  rq_init_comm_if_connected(9, "1")
  rq_init_comm_if_connected(2, "2")
  rq_init_comm_if_connected(3, "3")
  rq_init_comm_if_connected(4, "4")
  rq_print_connected_grippers()
  rq_gripper_communication_thread = run rq_gripper_communication()
  set_closed_norm(97.6470588235294, 1)
  set_open_norm(1.1764705882352942, 1)
  set_closed_mm(0.0, 1)
  set_open_mm(53.0, 1)
  set_closed_norm(100.0, 2)
  set_open_norm(0.0, 2)
  set_closed_mm(0.0, 2)
  set_open_mm(50.0, 2)
  set_closed_norm(100.0, 3)
  set_open_norm(0.0, 3)
  set_closed_mm(0.0, 3)
  set_open_mm(50.0, 3)
  set_closed_norm(100.0, 4)
  set_open_norm(0.0, 4)
  set_closed_mm(0.0, 4)
  set_open_mm(50.0, 4)
  rq_current_limit_enabled = False
  while(not rq_gripper_communication_thread_started):
      sync()
  end
  # end: URCap Installation Node
  global AMR_Position=struct(position_identifier=0, x1=0, x2=0, y1=0, y2=0, theta1=0, theta2=0)
  global CAM_Pose=p[0,0,0,0,0,0]
  global CAM_Relation=""
  global CMD_Abort=  False
  global CMD_Clear=  False
  global CMD_Reset=  False
  global CMD_Start=  False
  global CMD_Suspend=  False
  global CMD_Unhold=  False
  global CMD_Unsuspend=  False
  global CNT_Rack_Output=0
  global FNC_Freedrive=  False
  global PRC_TubCounter=0
  global PRC_TubNumber=0
  global STP=0
  global easyPickCount=0
  global easyPickCount_1=0
  global easyPickCount_2=0
  global easyPickCount_3=0
  global easyPickNoObj=0
  global easyPickNoObj_1=0
  global easyPickNoObj_2=0
  global easyPickNoObj_3=0
  global easyPickParts=0
  global easyPickParts_1=0
  global easyPickParts_2=0
  global easyPickParts_3=0
  global TMR_Barcode=0
  global Waypoint_6_p=p[.008800512419, -.547926542621, .402696567415, -.589884378425, -.007228654778, -.061268144704]
  global Waypoint_6_q=[-1.2044575850116175, -1.3416667741588135, -1.8272563219070435, -0.9884541195682068, 1.3621035814285278, -2.7712565104113978]
  global Waypoint_18_p=p[-.178371829612, -.433927395311, .368082383916, -.086593488055, .704679941724, -.007869906074]
  global Waypoint_18_q=[-1.265390698109762, -1.3355963987163086, -1.7944865226745605, -1.7402602634825648, 0.8780410885810852, -2.7713127771960657]
  global Waypoint_12_p=p[.008800512419, -.547926542621, .402696567415, -.589884378425, -.007228654778, -.061268144704]
  global Waypoint_12_q=[-1.2044575850116175, -1.3416667741588135, -1.8272563219070435, -0.9884541195682068, 1.3621035814285278, -2.7712565104113978]
  global Waypoint_19_p=p[-.178371829612, -.433927395311, .368082383916, -.086593488055, .704679941724, -.007869906074]
  global Waypoint_19_q=[-1.265390698109762, -1.3355963987163086, -1.7944865226745605, -1.7402602634825648, 0.8780410885810852, -2.7713127771960657]
  global Vial_above_p=p[.017105793010, -.652093028359, .184920586844, .000000000272, .000000000270, 1.564063451276]
  global Vial_above_q=[-1.3375440709712851, -1.9618096977868804, -1.4665759083780685, -1.2837941559171444, 1.5732503672317195, -4.47276330421513]
  global Vial_pick_point_p=p[.017105792852, -.648922724010, .093307568731, .000000000271, .000000000270, 1.564063451276]
  global Vial_pick_point_q=[-1.3366329456391917, -2.0375277831965413, -1.6071432798879028, -1.0675084332049813, 1.57309887265915, -4.471135348858068]
  global Waypoint_20_p=p[.019227646885, -.648669633640, .184920586950, .000000000000, .000000000000, .024063451426]
  global Waypoint_20_q=[-1.3331129109407733, -1.9540750545686123, -1.4775914902901128, -1.280581784992414, 1.5733500744865856, -2.928303704452631]
  global Waypoint_33_p=p[-.032361834699, -.348336136197, .391475576335, -.000008499254, .000014589902, -.004651426820]
  global Waypoint_33_q=[-1.2709335019096129, -1.1914598663441005, -1.708995335060501, -1.8117888533498316, 1.5729683532263925, -2.8379347397710237]
  global Vial_3FG_place_p=p[-.031858676359, -.349402499566, .145301120695, .000000000000, .000000000000, .000000000000]
  global Vial_3FG_place_q=[-1.2723975525801707, -1.252376585823825, -2.3128114007049496, -1.1470592278900167, 1.5730548099411423, -2.8414815174610535]
  global Waypoint_34_p=p[-.032361834699, -.348336136197, .391475576335, -.000008499254, .000014589902, -.004651426820]
  global Waypoint_34_q=[-1.2709335019096129, -1.1914598663441005, -1.708995335060501, -1.8117888533498316, 1.5729683532263925, -2.8379347397710237]
  global cap_dump_p=p[-.139168676487, -.420163541420, .146096395183, .000000000000, .000000000000, .000000000000]
  global cap_dump_q=[-1.584588644510994, -1.5093464179777323, -2.1118449369620347, -1.091059703602438, 1.5728943834877336, -3.154014906686923]
  global Waypoint_35_p=p[-.032361834699, -.348336136197, .391475576335, -.000008499254, .000014589902, -.004651426820]
  global Waypoint_35_q=[-1.2709335019096129, -1.1914598663441005, -1.708995335060501, -1.8117888533498316, 1.5729683532263925, -2.8379347397710237]
  global Waypoint_36_p=p[-.032361834699, -.348336136197, .391475576335, -.000008499254, .000014589902, -.004651426820]
  global Waypoint_36_q=[-1.2709335019096129, -1.1914598663441005, -1.708995335060501, -1.8117888533498316, 1.5729683532263925, -2.8379347397710237]
  global Waypoint_37_p=p[-.032361834699, -.348336136197, .391475576335, -.000008499254, .000014589902, -.004651426820]
  global Waypoint_37_q=[-1.2709335019096129, -1.1914598663441005, -1.708995335060501, -1.8117888533498316, 1.5729683532263925, -2.8379347397710237]
  global Vial_liq_above_p=p[-.025303660977, -.338758622354, .426628485936, -1.315858642253, .800043520260, -.928295855026]
  global Vial_liq_above_q=[-0.3789628187762659, -1.5149522957256814, -2.263045310974121, 0.7870649534412841, -0.750984017048971, -3.2237566153155726]
  global Vial_liq_pick_1_p=p[-.002660428945, -.335984893034, .159389832934, -1.150456778400, .673175527684, -1.010612657503]
  global Vial_liq_pick_1_q=[-0.3660772482501429, -1.4503649038127442, -2.4056053161621094, -1.994692941705221, 0.8039668202400208, -0.2508929411517542]
  global Vial_liq_pick_2_p=p[-.041402486291, -.356791603314, .125395323246, -1.143483969075, .651070210027, -.878721885453]
  global Vial_liq_pick_2_q=[-0.4426233705502476, -1.437252121513727, -2.551930962114307, -1.776528229806984, 0.6562026234073748, -0.43018811960029524]
  global Liquid_midway_p=p[.057575295009, -.583081747994, .306414980749, -1.351675548728, .120935756539, -.096908606303]
  global Liquid_midway_q=[-0.895174805318014, -1.7035466633238734, -2.380953073501587, 0.631549521083496, 0.7706599235534668, -2.9455552736865442]
  global shake_1_p=p[.057574880217, -.583085370269, .306422893466, -1.360996190983, -.155555042453, -.438136255921]
  global shake_1_q=[-0.8951800505267542, -1.7035466633238734, -2.380937099456787, 0.6315542894550782, 0.7706599235534669, -2.5394540616517496]
  global shake_2_p=p[.057581636113, -.583090570002, .306439684073, -1.308767904323, .368530312677, .214926493520]
  global shake_2_q=[-0.8951714674579065, -1.7035395107665003, -2.380906343460083, 0.6315504747578125, 0.7706480026245118, -3.3161255787892268]
  global drop_above_1_p=p[.268235025993, -.467784390499, .226219872376, -1.027832627524, -.430841408251, 1.004603115937]
  global drop_above_1_q=[-0.935645882283346, -1.6663371525206507, -2.4252893924713135, 0.41966931402172847, 1.8470635414123535, -3.4600217978106897]
  global drop_above_2_p=p[.219042229014, -.470775657081, .133754190740, -.313004595901, -.344395319364, 1.500564994056]
  global drop_above_2_q=[-1.0601594887284795, -1.70046459045642, -2.0799996233759863, -0.7243227230676759, 1.9429634314685202, -4.115129153870795]
  global liq_tran_1_p=p[.213067510942, -.469567035397, .100231043184, .251862243732, .217902579404, 1.592812335393]
  global liq_tran_1_q=[-0.7789645168037476, -1.822364827406652, -1.8643518410805573, -1.252158963840138, 1.3768134449520435, -3.9328333233290254]
  global Waypoint_21_p=p[.187119460405, -.493959476151, .133754190608, -.313004596540, -.344395317757, 1.500564993991]
  global Waypoint_21_q=[-1.1418328121400876, -1.7310553375189475, -2.033634768766424, -0.772026910513711, 1.958578934631971, -4.201588449364511]
  global liq_tran_2_p=p[.195957706507, -.493022614126, .100231042689, .160718757180, .109807038912, 1.525321508623]
  global liq_tran_2_q=[-0.881740380645474, -1.8244526267589851, -1.865100964490387, -1.1608866323693583, 1.4631433601076713, -3.973915130363038]
  global Vial_drop_above_p=p[.000324902251, -.648569523142, .221894115667, -.873462921366, 1.165852672573, -1.482720593185]
  global Vial_drop_above_q=[-1.0576906334721352, -2.393016994184633, -0.9236232851859159, -2.5729213042279273, 0.7903331288549689, -0.33286325848155585]
  global Vial_liq_drop_p=p[.001020867953, -.647659915585, .092915870838, -.834762611599, 1.081942994823, -1.540647900176]
  global Vial_liq_drop_q=[-1.0631954168193474, -2.4447642951220825, -1.128811017825127, -2.1983115491972294, 0.8130148661460634, -0.38984988696911316]
  global Waypoint_9_p=p[.206300564882, -.401796282405, .209941275233, .000000000049, .000000000063, 1.560839127857]
  global Waypoint_9_q=[-0.7963359454512808, -1.4686025034365713, -1.9726632321075135, -1.2709582822971974, 1.5730203818053559, -3.9272300959189193]
  global Waypoint_10_p=p[.200865824304, -.400817692024, .105072686738, .000000000049, .000000000061, 1.560839127855]
  global Waypoint_10_q=[-0.8042914374275529, -1.5824702465090397, -2.1630314773482997, -0.9667217216455377, 1.5726337265768082, -3.9342465798801403]
  global Waypoint_11_p=p[.200865824280, -.400817691999, .325177251663, .000000000049, .000000000061, 1.560839127855]
  global Waypoint_11_q=[-0.8031609769098491, -1.4190566846320642, -1.7173307870816634, -1.5758364190022327, 1.5730457436482617, -3.935202548332848]
  global Waypoint_7_p=p[-.615828862681, .233809157513, .299999999960, .005115849907, .008741794022, -2.111813105778]
  global Waypoint_7_q=[-3.2957401409809868, -1.9361965884744503, -1.2056078493731617, -1.569266158150004, 1.5650998100608482, -2.7562028470627613]
  global Waypoint_8_p=p[-.615828862366, .233809157463, .013910424379, .005115849905, .008741794020, -2.111813105780]
  global Waypoint_8_q=[-3.2964782505943173, -2.1586184138220776, -1.6500090431308791, -0.9024541777239836, 1.5648120752692236, -2.7547026290098384]
  global Container_midwa_p=p[-.379239199143, -.127191311915, .299999999998, .000000000046, -.000000000021, -1.247199999994]
  global Container_midwa_q=[-2.477408934449926, -1.2969853503591224, -1.875639182904262, -1.539621866126728, 1.5731943360401213, -2.8009955944022717]
  global Container_capt_p=p[-.525590029047, .407247642794, .411588185841, -.000000000107, .000000000065, -2.896148821900]
  global Container_capt_q=[-3.5968351615224767, -2.0050156108707204, -0.8176271154495112, -1.8895759482008394, 1.5730967555598792, -2.2743681102957645]
  global Waypoint_13_p=p[-.479450777041, .284140798427, .125270103493, -.276792173670, 2.098433187455, -2.121256516887]
  global Waypoint_13_q=[-2.8915050665484827, -1.9549266300597132, -2.2318272590637207, -1.6654960117735804, 0.020810842514038086, -0.4019392172442835]
  global Waypoint_1_p=p[-.472820924464, .292439826304, .207418370234, -.259787347864, -2.053484648504, 2.070709755662]
  global Waypoint_1_q=[-2.969927421603815, -2.07168115810532, -1.6835546062719366, -2.4953958198513964, 0.4489790927922641, -0.005578998612037367]
  global Waypoint_2_p=p[-.312961047461, -.152991312519, .223609826854, -.745314530454, -1.713873240489, 1.673341715282]
  global Waypoint_2_q=[-2.3560472170459192, -2.183784624139303, -1.4583134651184082, -2.6435262165465296, 1.6522362232208252, 0.043451953679323196]
  global Waypoint_3_p=p[-.113749865836, -.390110151572, .317307487562, -.519383711706, -.839884211339, 1.756868173041]
  global Waypoint_3_q=[-1.8909733931170862, -1.720626016656393, -1.5115610361099243, -2.1240560017027796, 2.1809096336364746, 0.7227501273155212]
  global Waypoint_15_p=p[.029144035010, -.436802470887, .327885032028, -.521560953301, -.623641814548, 1.862659450154]
  global Waypoint_15_q=[-1.564817253743307, -1.556895188321807, -1.6826975345611572, -1.6944714985289515, 2.2362685203552246, 1.117417335510254]
  global Waypoint_14_p=p[.068712235638, -.569419545175, .285215357659, -.679242949116, -.712065334485, 1.394044574094]
  global Waypoint_14_q=[-1.5731792953485346, -1.8029235103747094, -1.6781008808776736, -1.2218450646111982, 2.4719572998240125, 1.6394218026856375]
  global Waypoint_4_p=p[-.047220457210, -.557624911767, .136370962514, -.679242949107, -.712065334475, 1.394044574096]
  global Waypoint_4_q=[-1.7740079055958748, -2.0023561428872334, -1.7577251142892676, -1.18903287716154, 2.4487287370345143, 1.322902469273079]
  global Waypoint_25_p=p[.065436479647, -.569388431626, .287820755049, -.679242949185, -.712065334557, 1.394044574070]
  global Waypoint_25_q=[-1.5789263550890595, -1.8020194754825436, -1.6702557537748035, -1.237882536889547, 2.471995808083492, 1.6301087487321393]
  global Waypoint_16_p=p[-.389004373533, .141378246032, .266753254334, .000138837765, -.000085501467, -2.896077186553]
  global Waypoint_16_q=[-3.161701420154333, -1.339999469068478, -1.9293121603919792, -1.4429740688031423, 1.5733018961609508, -1.8361050683902924]
  global Waypoint_17_p=p[-.035033829322, -.360271411898, .346670090250, .000134865440, .000045012632, -1.419458520241]
  global Waypoint_17_q=[-1.2895553551337002, -1.2030299897931318, -1.8182548744695417, -1.6909649895170915, 1.5732755303988695, -1.4412981698552478]
  global Waypoint_22_p=p[-.031770714526, -.348511954549, .220918238016, .000139161477, .000025856264, -1.196413611588]
  global Waypoint_22_q=[-1.2709487693936374, -1.1814333631236558, -2.1531395672900686, -1.3776934646498997, 1.5734173079341525, -1.6444054353326152]
  global Waypoint_23_p=p[-.031891260245, -.348193352375, .178713903582, .000139161477, .000025856264, -1.196413611588]
  global Waypoint_23_q=[-1.271310670462512, -1.2113466935832626, -2.2466531062742767, -1.2542663946277255, 1.5733351685360857, -1.6443240949325606]
  global Waypoint_24_p=p[-.031773196918, -.348519672341, .270996689483, .000139161478, .000025856264, -1.196413611588]
  global Waypoint_24_q=[-1.270577047002206, -1.1645624227804543, -2.0341633523498315, -1.513540880628252, 1.5734258150982026, -1.6445600267865252]
  global Waypoint_26_p=p[-.030182364204, -.347335556538, .210997748016, .000000000000, .000000000000, .000000000000]
  global Waypoint_26_q=[-1.2651221433650806, -1.1831852705229569, -2.1779499233587867, -1.3511120827722447, 1.5732559871804586, -2.834886496531558]
  global Waypoint_27_p=p[-.030361452661, -.347415235983, .279538636214, -.000011913493, .000041085949, -.000383030923]
  global Waypoint_27_q=[-1.2651616254632172, -1.160029050867486, -2.014957410251413, -1.537262165299773, 1.573226049428862, -2.835263580680065]
  global Waypoint_28_p=p[-.154725436156, -.473256970882, .246188866975, -.000011913493, .000041085951, -.000383030922]
  global Waypoint_28_q=[-1.6148878344468836, -1.561261107922114, -1.7903420597774975, -1.3606341597365077, 1.5730936011867385, -3.1851320724005863]
  global Waypoint_29_p=p[-.145695304927, -.485909140058, .046677498463, -.000011913493, .000041085952, -.000383030922]
  global Waypoint_29_q=[-1.5959977509619323, -1.81576344419621, -2.079448728928398, -0.8170257869513264, 1.572443153678545, -3.1647042569483315]
  global Waypoint_38_p=p[-.145695304919, -.485909139930, .261430070956, -.000011913492, .000041085950, -.000383030921]
  global Waypoint_38_q=[-1.595239081389626, -1.5772455407988337, -1.734838265427694, -1.4001543934186973, 1.5731079270966675, -3.1656816807751103]
  global Waypoint_30_p=p[-.030182364221, -.347335556548, .265578332256, .000000000000, .000000000000, .000000000000]
  global Waypoint_30_q=[-1.2647056875423734, -1.1616486920426157, -2.0496625730758256, -1.500936273978276, 1.573279507668392, -2.8350442023705362]
  global Waypoint_31_p=p[-.030182364236, -.347335556501, .175832814209, .000000000000, .000000000000, .000000000000]
  global Waypoint_31_q=[-1.2653656161933107, -1.210901321223588, -2.254656599340546, -1.2466892005088948, 1.573177712256868, -2.834760980417842]
  global Waypoint_32_p=p[-.030182364238, -.347335556494, .316066543581, .000000000000, .000000000000, .000000000000]
  global Waypoint_32_q=[-1.2642809742958807, -1.161008069550718, -1.9212694317539043, -1.629970222817029, 1.5732134180415143, -2.835147596020935]
  global Waypoint_39_p=p[.137772150180, -.577759956854, .299999999946, .000000000217, -.000000000207, -1.594351842625]
  global Waypoint_39_q=[-1.108978697428574, -1.776486680444405, -1.413737665315093, -1.5218908901738937, 1.5733062372356947, -1.0863866394180182]
  global Waypoint_41_p=p[.074222967010, -.565641640647, .234620140366, -.516884386806, .529223682286, -1.529619060506]
  global Waypoint_41_q=[-0.9596722604286052, -1.8767069964135548, -1.4892746174057256, -1.7813862040292285, 1.0520698599867686, -0.8199687448260349]
  global Waypoint_40_p=p[.039987741677, -.564832865048, .191055405868, -.767560686167, .343136533060, -2.241315728308]
  global Waypoint_40_q=[-1.0070649180116558, -1.8745927522477324, -1.6139175023195245, -1.6337474788493545, 1.032708081143138, -0.11587278312988403]
  global Waypoint_42_p=p[.041363380882, -.564865360786, .192805844739, .278500165520, .624117100927, .762272396553]
  global Waypoint_42_q=[-1.0050718976263102, -1.8744386685524779, -1.609151451954446, -1.6399653140247947, 1.0334006002355505, -3.254032861659603]
  global Waypoint_43_p=p[.041363380884, -.564865360793, .192805844731, .973435683493, .064103649514, 2.808306925555]
  global Waypoint_43_q=[-1.0050547674917611, -1.8743226123411425, -1.6093213313885109, -1.6397178529514314, 1.0333615331919874, -5.424787697362414]
  global Waypoint_44_p=p[.040882892233, -.564854254876, .192193763716, .110913882012, .659173708659, .275719738520]
  global Waypoint_44_q=[-1.0057704811530535, -1.8745207681598055, -1.6107765025572558, -1.637858394640876, 1.033164860873599, -2.7487836132940755]
  global Waypoint_45_p=p[.042647731639, -.564895808997, .194439423694, -.451694728506, .563172064821, -1.343350300184]
  global Waypoint_45_q=[-1.0032860829914387, -1.8741561795270565, -1.6048483308761785, -1.6453689714776623, 1.0342050634514657, -1.06078829880322]
  global Waypoint_46_p=p[.099944144487, -.566244126804, .267342790130, -.451694834765, .563172023386, -1.343350532536]
  global Waypoint_46_q=[-0.9257438092434924, -1.889970530402497, -1.3828165217629076, -1.8916791100652528, 1.0664350961373816, -0.9805910833329659]
  global Waypoint_47_p=p[.099944144444, -.566244126727, .267342790273, -.101742139519, .058679218003, -1.457888523314]
  global Waypoint_47_q=[-1.1112623176383014, -1.729989471869196, -1.5530029871033957, -1.4442770617454777, 1.4670579052775654, -1.2224020460061675]
  global Waypoint_48_p=p[-.136182767566, -.647487115908, .294247768372, -.101742139549, .058679218020, -1.457888523312]
  global Waypoint_48_q=[-1.532196177857717, -1.9115932455375173, -1.2651848069729779, -1.5055651746702665, 1.4703193777418382, -1.646379689188814]
  global Waypoint_49_p=p[-.159024328559, -.641021381179, .047691706070, -.000000000033, -.000000000027, -1.457897102937]
  global Waypoint_49_q=[-1.6098490079965062, -2.1164987141784586, -1.6156631902166785, -0.9800092198841526, 1.573231151532669, -1.722204302767242]
  global Waypoint_50_p=p[-.159024328558, -.641021381151, .291114489351, -.000000000033, -.000000000027, -1.457897102937]
  global Waypoint_50_q=[-1.609190265995684, -1.9426985888940234, -1.2189094859258596, -1.55056435122874, 1.5734384912955113, -1.7235116759964022]
  global Waypoint_51_p=p[-.138513366863, -.390317608895, .390026797065, .985058163405, .076630161240, 2.827313005358]
  global Waypoint_51_q=[-1.1615256227675719, -1.2926165506592575, -1.7164354353247306, -2.007781815499934, 0.9660985548762523, 0.6591122264722848]
  global Waypoint_52_p=p[.200663338988, -.570117491939, .330074050008, 1.360500824927, .021700159056, 2.681649888904]
  global Waypoint_52_q=[-0.766974602501266, -2.1699046207818107, -0.8659485470448569, -2.4759404440644786, 1.0197680658968387, 1.1887972982227069]
  global Waypoint_53_p=p[.200650292861, -.570238752026, .330084459991, 1.360500825815, .021700154388, 2.681649888469]
  global Waypoint_53_q=[-0.7671117850166942, -2.170180210127774, -0.8654875324671831, -2.4760661058854714, 1.019668964673781, 1.1886838746103445]
  global Waypoint_54_p=p[.143029822311, -.569853361759, .275754213782, 1.297896664289, .026410127072, 2.712872144875]
  global Waypoint_54_q=[-0.8339941389801577, -2.0499669090260237, -1.181859109742545, -2.1992567984298894, 0.9933974691724003, 1.1053015960835664]
  global Waypoint_55_p=p[.073857253409, -.577012553496, .221504790513, 1.297896665457, .026410123899, 2.712872144362]
  global Waypoint_55_q=[-0.9235026509638331, -2.0031911550113533, -1.4013130080059835, -1.9791459123699324, 0.9364696407276547, 1.0224867664664226]
  global Waypoint_56_p=p[.135677267144, -.579447716527, .242231366835, 1.555421348248, .015405426287, 2.555899922373]
  global Waypoint_56_q=[-0.8277598345563266, -2.1783820448240228, -1.1390951780517948, -2.3437042464770936, 0.9222576608739947, 1.2572681804986878]
  global Waypoint_57_p=p[.143391004007, -.581808738942, .226065325532, 1.639743959545, .007914821713, 2.502360786858]
  global Waypoint_57_q=[-0.8163397121067408, -2.2409861865625498, -1.1056400409378426, -2.4000192569642436, 0.9131014133193622, 1.3141118037187605]
  global Waypoint_59_p=p[.272401132286, -.578182925380, .239561357365, 2.126997331910, .113921148153, 2.155615020515]
  global Waypoint_59_q=[-0.6600120703326624, -2.700596948663229, -0.4450863301753998, -3.1158048115172328, 0.9327830672264099, 1.686402678489685]
  global Waypoint_58_p=p[.223648508176, -.578477552733, .276546452136, 2.174288010107, -.044108754041, 2.058653287678]
  global Waypoint_58_q=[-0.7290484882560344, -2.6749849159411134, -0.44426632073579775, -3.220833992584847, 0.9665895014735898, 1.686536774549042]
  global Waypoint_60_p=p[-.013316432876, -.544772031582, .383371643081, 2.208233379808, .037543335712, 2.097559881761]
  global Waypoint_60_q=[-0.9328326161883087, -2.0999933666355775, -1.1958015693111372, -3.060905141293654, 0.690378518537611, 1.7121940951337198]
  global Waypoint_61_p=p[-.412188693372, -.356446875193, .383371643081, 1.751740964455, -.739956256289, 1.600691174920]
  global Waypoint_61_q=[-1.766185342973321, -2.0999933666355775, -1.1958015693111372, -3.060905141293654, 0.690378518537611, 1.7121940951337198]
  global Waypoint_62_p=p[-.542658707241, -.114281911009, .251261544113, 1.813043609523, -.679411528034, 1.655271622964]
  global Waypoint_62_q=[-2.158300033470912, -1.9418836862428677, -1.8142999147147894, -2.778920736683023, 0.21900622104017292, 1.8983390235012934]
  global Waypoint_63_p=p[-.532496162227, -.127810170801, .159342327524, 1.813043609478, -.679411528027, 1.655271622994]
  global Waypoint_63_q=[-2.1232624524640213, -2.086114053133292, -1.8911847933380095, -2.5248779786918614, 0.2536249317365024, 1.864405460969639]
  global Waypoint_64_p=p[-.576034890047, -.066269986912, .306739617770, .862065193359, -.255405331227, 2.195240951653]
  global Waypoint_64_q=[-2.4808268779922003, -1.5303848711262056, -1.876845562237385, -1.1257011427858359, 0.8740163290385958, -0.15002503295170655]
  global Waypoint_65_p=p[-.581965326699, -.059291422286, .312082125679, .862065195757, -.255405329473, 2.195240950921]
  global Waypoint_65_q=[-2.500621389999687, -1.5361955180345959, -1.8614018767844556, -1.1190332887072278, 0.8777181708365909, -0.17540933674578696]
  global Waypoint_66_p=p[-.581965326670, -.059291422265, .290575803625, .862065195756, -.255405329472, 2.195240950921]
  global Waypoint_66_q=[-2.5007210652259566, -1.5510704265538795, -1.9040561970342402, -1.0615823481403304, 0.8776641555740685, -0.17528706367848557]
  global Waypoint_67_p=p[-.581965326627, -.059291422244, .350142125738, 1.757497900770, -.677813691618, 1.696469016977]
  global Waypoint_67_q=[-2.3014470577960933, -1.774776476208789, -1.7081605706825291, -2.8433626113276596, 0.07508598567825443, 1.682946898281932]
  global Waypoint_68_p=p[-.333292906431, -.480744165508, .350142125738, 2.217519979286, .140864133573, 2.209123277630]
  global Waypoint_68_q=[-1.438387057796029, -1.774776476208789, -1.7081605706825291, -2.8433626113276596, 0.07508598567825443, 1.682946898281932]
  global TMR_Barcode_is_counting=False
  thread Timer_Thread():
    while (True):
      if (TMR_Barcode_is_counting):
        TMR_Barcode = TMR_Barcode + get_steptime()
      end
      sync()
    end
  end
  run Timer_Thread()
  def Sub_Vision_V18():
    $ 882 "Sub_Vision_V18" "noBreak"
    $ 883 "PreSettings"
    $ 884 "CAM_LM_Detected≔ False "
    global CAM_LM_Detected=  False
    $ 885 "CAM_Captures≔0"
    global CAM_Captures=0
    $ 886 "CAM_Pose≔p[0,0,0,0,0,0]"
    global CAM_Pose=p[0,0,0,0,0,0]
    $ 887 "CAM_LM_Refinmnt≔ False "
    global CAM_LM_Refinmnt=  False
    $ 888 "CAM_LM_Refined≔ False "
    global CAM_LM_Refined=  False
    $ 889 "CAM_LM_Deviatn≔p[0,0,0,0,0,0]"
    global CAM_LM_Deviatn=p[0,0,0,0,0,0]
    $ 890 "CAM_LM_ID≔0"
    global CAM_LM_ID=0
    $ 891 "CAM_Done≔ False "
    global CAM_Done=  False
    $ 892 "CAM_CNT_Obj≔0"
    global CAM_CNT_Obj=0
    $ 893 "CAM_Result = []"
    CAM_Result = []
    $ 894 "OBJ_Detected≔ False "
    global OBJ_Detected=  False
    $ 895 "FRM_Reference≔p[0,0,0,0,0,0]"
    global FRM_Reference=p[0,0,0,0,0,0]
    $ 896 "'=========='"
    # '=========='
    $ 897 "Switch Action"
    switch_1 = Action
    $ 898 "Case 13"
    if (13 == switch_1):
    elif (15 == switch_1):
      $ 1016 "Case 15"
    elif (131 == switch_1):
      $ 1062 "Case 131"
      $ 1063 "Read (SensoPart)"
      $ 1064 "Action_Info≔'search for landmark'"
      global Action_Info="search for landmark"
      $ 1065 "CAM_LM≔CAM_LMs[4]"
      global CAM_LM=CAM_LMs[4]
      $ 1066 "CAM_Relation≔CAM_LM.capture_relation"
      global CAM_Relation=CAM_LM.capture_relation
      $ 1067 "go to capture pose"
      $ 1070 "If ITM_ID≟1 and JIG≟7"
      if (ITM_ID == 1  and  JIG == 7):
        $ 1071 "PSE_T≔uLM_Cap_SSRack"
        global PSE_T=uLM_Cap_SSRack
      else:
        $ 1072 "ElseIf ITM_ID≟5 and JIG≟7"
        if (ITM_ID == 5  and  JIG == 7):
          $ 1073 "PSE_T≔FRM_Cap_SSRack"
          global PSE_T=FRM_Cap_SSRack
        else:
          $ 1074 "ElseIf ITM_ID≟13 and JIG≟7"
          if (ITM_ID == 13  and  JIG == 7):
            $ 1075 "PSE_T≔FRM_pick_rack_const"
            global PSE_T=p[-0.5568395192387274,0.34423986364170267,0.44698620470146266,-1.0069110132199915E-6,3.378712467497258E-5,-8.002029546773325E-6]
          end
        end
      end
      $ 1076 "do_transition(PSE_T, keep_rxry=False)"
      do_transition(PSE_T, keep_rxry=False)
      $ 1077 "Set"
      set_tcp(p[0.0,0.0,0.161,3.1415,0.0,0.0])
      $ 1078 "MoveJ"
      $ 1079 "PSE_T" "breakAfter"
      movej(PSE_T, a=1.3962634015954636, v=1.7453292519943295)
      $ 1080 "CAM_Pose≔get_actual_tcp_pose()"
      global CAM_Pose= get_actual_tcp_pose ()
      $ 1081 "Loop  not CAM_Done and  not ERROR.FLAG and  not CMD_Stop"
      while (  not  CAM_Done  and    not  ERROR.FLAG  and    not  CMD_Stop):
        $ 1082 "adjust capture pose"
        $ 1083 "If CAM_LM_Detected and CAM_LM_Refinmnt"
        if (CAM_LM_Detected  and  CAM_LM_Refinmnt):
          $ 1084 "PSE_T≔p[0,0,0.300,0,0,0]"
          global PSE_T=p[0,0,0.300,0,0,0]
          $ 1085 "CAM_Pose≔PSE_T"
          global CAM_Pose=PSE_T
          $ 1086 "If  not is_reachable(FRM_Reference,[PSE_T])"
          if (  not  is_reachable(FRM_Reference,[PSE_T])):
            $ 1087 "Error"
            $ 1088 "set_error(ERROR_POSE_NOT_REACHABLE)"
            set_error(ERROR_POSE_NOT_REACHABLE)
          end
          $ 1089 "If  not ERROR.FLAG"
          if (  not  ERROR.FLAG):
            $ 1090 "MoveJ"
            $ 1091 "PSE_T" "breakAfter"
            set_tcp(p[0.0,0.0,0.161,0.0,0.0,0.0])
            movej(pose_trans(FRM_Reference, PSE_T), a=0.8726646259971648, v=1.3962634015954636)
            $ 1092 "CAM_LM_Refined≔ True "
            global CAM_LM_Refined=  True
          end
        else:
          $ 1093 "ElseIf  not CAM_LM_Detected and CAM_Captures>0"
          if (  not  CAM_LM_Detected  and  CAM_Captures>0):
            $ 1094 "MoveL"
            $ 1095 "If FRM_Reference≟p[0,0,0,0,0,0]"
            if (FRM_Reference == p[0,0,0,0,0,0]):
              $ 1096 "PSE_T≔get_random_pose(pose_ref=CAM_Pose, mode='cubic', range_max=[0.150,0.150,0.015])"
              global PSE_T=get_random_pose(pose_ref=CAM_Pose, mode="cubic", range_max=[0.150,0.150,0.015])
            else:
              $ 1101 "Else" "noBreak"
              $ 1102 "PSE_T≔get_random_pose(pose_ref=CAM_Pose, mode='rotation', range_max=[10,10,0])"
              global PSE_T=get_random_pose(pose_ref=CAM_Pose, mode="rotation", range_max=[10,10,0])
              $ 1103 "CAM_LM_Refined≔ True "
              global CAM_LM_Refined=  True
            end
            $ 1104 "If get_inverse_kin_has_solution(pose_trans(FRM_Reference, PSE_T))"
            if (get_inverse_kin_has_solution( pose_trans (FRM_Reference, PSE_T))):
              $ 1105 "Comment"
              # Comment
              $ 1106 "PSE_T" "breakAfter"
              set_tcp(p[0.0,0.0,0.161,3.1415,0.0,0.0])
              movel(pose_trans(FRM_Reference, PSE_T), a=0.03, v=0.05)
            else:
              $ 1107 "Else" "noBreak"
              $ 1108 "'If random pose is out of reach, set the initial cam pose'"
              # 'If random pose is out of reach, set the initial cam pose'
              $ 1109 "PSE_T≔CAM_Pose"
              global PSE_T=CAM_Pose
            end
          end
        end
        $ 1110 "Wait: 2.0"
        sleep(2.0)
        $ 1111 "trigger"
        # begin: URCap Program Node
        #   Source: SensoPart VISOR Robotic, 2.0.0, SensoPart Industriesensorik GmbH
        #   Type: VISOR Trigger
        $ 1112 "# 1 VISOR Trigger"
        visor_changeJob(1, "Landmark_INVITE_2", 6000)
        visor_trigger(1, 6000, "arm")
        # end: URCap Program Node
        $ 1116 "TM_3D_Found≔visor_partsFound(1)"
        global TM_3D_Found= visor_partsFound (1)
        $ 1117 "If TM_3D_Found>0"
        if (TM_3D_Found>0):
          $ 1118 "CAM_LM_Detected≔ True "
          global CAM_LM_Detected=  True
          $ 1119 "CAM_Captures≔0"
          global CAM_Captures=0
        else:
          $ 1120 "Else" "noBreak"
          $ 1121 "CAM_LM_Detected≔ False "
          global CAM_LM_Detected=  False
          $ 1122 "CAM_Captures≔CAM_Captures+1"
          global CAM_Captures=CAM_Captures+1
        end
        $ 1127 "result"
        $ 1128 "If CAM_LM_Detected"
        if (CAM_LM_Detected):
          $ 1129 "If (CAM_LM_Refinmnt and CAM_LM_Refined) or  not CAM_LM_Refinmnt"
          if ((CAM_LM_Refinmnt  and  CAM_LM_Refined)  or    not  CAM_LM_Refinmnt):
            $ 1187 "If ITM_ID≟1 and JIG≟7"
            if (ITM_ID == 1  and  JIG == 7):
              $ 1188 "CAM_LM_SSRack≔visor_getPose3d(1, 0)"
              global CAM_LM_SSRack= visor_getPose3d (1, 0)
            else:
              $ 1189 "ElseIf ITM_ID≟5 and JIG≟7"
              if (ITM_ID == 5  and  JIG == 7):
                $ 1190 "CAM_LM_SSRack≔visor_getPose3d(1, 0)"
                global CAM_LM_SSRack= visor_getPose3d (1, 0)
              else:
                $ 1191 "ElseIf ITM_ID≟13 and JIG≟7"
                if (ITM_ID == 13  and  JIG == 7):
                  $ 1192 "CAM_LM_Bott≔visor_getPose3d(1, 0)"
                  global CAM_LM_Bott= visor_getPose3d (1, 0)
                end
              end
            end
            $ 1193 "CAM_Done≔ True "
            global CAM_Done=  True
          end
        else:
          $ 1194 "ElseIf  not CAM_LM_Detected and CAM_Captures<CAM_PRM_Retries"
          if (  not  CAM_LM_Detected  and  CAM_Captures<CAM_PRM_Retries):
            $ 1195 "CAM_LM_Refined≔ False "
            global CAM_LM_Refined=  False
          else:
            $ 1196 "ElseIf CAM_Captures≥CAM_PRM_Retries"
            if (CAM_Captures >= CAM_PRM_Retries):
              $ 1197 "CAM_Done≔ True "
              global CAM_Done=  True
              $ 1198 "Error"
              $ 1199 "set_error(ERROR_NO_LANDMARK)"
              set_error(ERROR_NO_LANDMARK)
            end
          end
        end
      end
    elif (151 == switch_1):
      $ 1200 "Case 151"
      $ 1201 "Detect (SensoPart)"
      $ 1202 "go to capture pose"
      $ 1203 "FRM_Reference≔FRM_Cap_SSRack"
      global FRM_Reference=FRM_Cap_SSRack
      $ 1204 "PSE_T≔p[0,0,-0.00,0,0,0]"
      global PSE_T=p[0,0,-0.00,0,0,0]
      $ 1205 "do_transition(pose_trans(FRM_Reference, PSE_T), keep_rxry=False)"
      do_transition( pose_trans (FRM_Reference, PSE_T), keep_rxry=False)
      $ 1206 "JNT_Q≔get_actual_joint_positions()"
      global JNT_Q= get_actual_joint_positions ()
      $ 1207 "JNT_Q≔[JNT_Q[0], JNT_Q[1], JNT_Q[2], JNT_Q[3], JNT_Q[4], 0]"
      global JNT_Q=[JNT_Q[0], JNT_Q[1], JNT_Q[2], JNT_Q[3], JNT_Q[4], 0]
      $ 1208 "Set"
      set_tcp(p[0.0,0.0,0.161,3.1415,0.0,0.0])
      $ 1209 "movej(get_inverse_kin(pose_trans(FRM_Reference, PSE_T), qnear=JNT_Q))"
      movej(get_inverse_kin( pose_trans (FRM_Reference, PSE_T), qnear=JNT_Q))
      $ 1210 "CAM_Pose≔pose_trans(pose_inv(FRM_Reference), get_actual_tcp_pose())"
      global CAM_Pose= pose_trans ( pose_inv (FRM_Reference),  get_actual_tcp_pose ())
      $ 1211 "Loop  not CAM_Done and  not ERROR.FLAG and  not CMD_Stop"
      while (  not  CAM_Done  and    not  ERROR.FLAG  and    not  CMD_Stop):
        $ 1212 "If  not OBJ_Detected and CAM_Captures>0"
        if (  not  OBJ_Detected  and  CAM_Captures>0):
          $ 1213 "MoveL"
          $ 1214 "If FRM_Reference≟p[0,0,0,0,0,0]"
          if (FRM_Reference == p[0,0,0,0,0,0]):
            $ 1216 "PSE_T≔get_random_pose(pose_ref=CAM_Pose, mode='rotation', range_max=[15,15,0])"
            global PSE_T=get_random_pose(pose_ref=CAM_Pose, mode="rotation", range_max=[15,15,0])
          else:
            $ 1217 "Else" "noBreak"
            $ 1218 "PSE_T≔get_random_pose(pose_ref=CAM_Pose, mode='rotation', range_max=[10,10,0])"
            global PSE_T=get_random_pose(pose_ref=CAM_Pose, mode="rotation", range_max=[10,10,0])
          end
          $ 1219 "If get_inverse_kin_has_solution(pose_trans(FRM_Reference, PSE_T))"
          if (get_inverse_kin_has_solution( pose_trans (FRM_Reference, PSE_T))):
            $ 1220 "PSE_T" "breakAfter"
            set_tcp(p[0.0,0.0,0.161,3.1415,0.0,0.0])
            movel(pose_trans(FRM_Reference, PSE_T), a=0.03, v=0.05)
          else:
            $ 1221 "Else" "noBreak"
            $ 1222 "'If random pose is out of reach, set the initial cam pose'"
            # 'If random pose is out of reach, set the initial cam pose'
            $ 1223 "PSE_T≔CAM_Pose"
            global PSE_T=CAM_Pose
            $ 1224 "PSE_T" "breakAfter"
            set_tcp(p[0.0,0.0,0.161,3.1415,0.0,0.0])
            movel(pose_trans(FRM_Reference, PSE_T), a=0.03, v=0.05)
          end
        end
        $ 1225 "Wait: 0.5"
        sleep(0.5)
        $ 1226 "Set"
        set_tcp(p[0.0,0.0,0.161,3.1415,0.0,0.0])
        # begin: URCap Program Node
        #   Source: SensoPart VISOR Robotic, 2.0.0, SensoPart Industriesensorik GmbH
        #   Type: VISOR Trigger
        $ 1227 "# 1 VISOR Trigger"
        visor_changeJob(1, "Object Detection Single", 6000)
        visor_trigger(1, 6000, "arm")
        # end: URCap Program Node
        $ 1228 "If visor_isResponseOk(1)"
        if ( visor_isResponseOk (1)):
          $ 1229 "CAM_CNT_Obj≔visor_partsFound(1)"
          global CAM_CNT_Obj= visor_partsFound (1)
          $ 1230 "CAM_OBJ_Pose≔visor_getPose3d(1, 0)"
          global CAM_OBJ_Pose= visor_getPose3d (1, 0)
          $ 1231 "If CAM_CNT_Obj>0"
          if (CAM_CNT_Obj>0):
            $ 1232 "CAM_OBJ_Color≔visor_getAdditionalData(1, 0)"
            global CAM_OBJ_Color= visor_getAdditionalData (1, 0)
            $ 1233 "CAM_DetectScore≔to_num(visor_getAdditionalData(1, 1))/1000"
            global CAM_DetectScore=to_num( visor_getAdditionalData (1, 1))/1000
            $ 1234 "OBJ_Detected≔ True "
            global OBJ_Detected=  True
          end
        else:
          $ 1235 "Else" "noBreak"
          $ 1236 "CAM_Captures≔CAM_Captures+1"
          global CAM_Captures=CAM_Captures+1
        end
        $ 1237 "If OBJ_Detected"
        if (OBJ_Detected):
          $ 1238 "Get object data"
          $ 1239 "PRC_CntDetect≔0"
          global PRC_CntDetect=0
          $ 1240 "Loop PRC_CntDetect<CAM_CNT_Obj"
          while (PRC_CntDetect<CAM_CNT_Obj):
            $ 1241 "get object and jig number"
            $ 1242 "If ITM_ID≟1 and JIG≟7"
            if (ITM_ID == 1  and  JIG == 7):
              $ 1243 "FRM_Reference≔FRM_Cap_SSRack"
              global FRM_Reference=FRM_Cap_SSRack
            else:
              $ 1244 "ElseIf ITM_ID≟5 and JIG≟7"
              if (ITM_ID == 5  and  JIG == 7):
                $ 1245 "FRM_Reference≔uLM_Cap_SSRack"
                global FRM_Reference=uLM_Cap_SSRack
              end
            end
            $ 1248 "PSE_T≔pose_trans(pose_inv(FRM_Reference), CAM_OBJ_Pose)"
            global PSE_T= pose_trans ( pose_inv (FRM_Reference), CAM_OBJ_Pose)
            $ 1249 "CAM_Result.append(get_pattern_counter(PSE_T, 'X', pattern=[10, 5], patternsize=[0.181, 0.081]))"
            CAM_Result.append(get_pattern_counter(PSE_T, "X", pattern=[10, 5], patternsize=[0.181, 0.081]))
            $ 1250 "PRC_CntDetect≔PRC_CntDetect+1"
            global PRC_CntDetect=PRC_CntDetect+1
          end
          $ 1251 "CAM_Done≔ True "
          global CAM_Done=  True
        else:
          $ 1252 "ElseIf CAM_Captures≥CAM_PRM_Retries"
          if (CAM_Captures >= CAM_PRM_Retries):
            $ 1253 "CAM_Done≔ True "
            global CAM_Done=  True
          else:
            $ 1254 "Else" "noBreak"
            $ 1255 "CAM_Captures≔CAM_Captures+1"
            global CAM_Captures=CAM_Captures+1
          end
        end
      end
    end
    $ 1256 "'=========='"
    # '=========='
    $ 1257 "PostSettings"
    $ 1258 "FRM_Reference≔p[0,0,0,0,0,0]"
    global FRM_Reference=p[0,0,0,0,0,0]
    $ 1259 "Set"
    set_tcp(p[0.0,0.0,0.161,3.1415,0.0,0.0])
    $ 1260 "CAM_Pose≔p[0,0,0,0,0,0]"
    global CAM_Pose=p[0,0,0,0,0,0]
    $ 1261 "Action≔0"
    global Action=0
    $ 1262 "Action_Info≔''"
    global Action_Info=""
  end
  def Sub_AMR_MiR_V3():
    $ 1263 "Sub_AMR_MiR_V3" "noBreak"
    $ 1264 "PreSettings"
    $ 1265 "AMR_TargetList≔[1,2,3,4,5,21,22,23,24,31,32,33,34,35,36,37,38,41]"
    global AMR_TargetList=[1,2,3,4,5,21,22,23,24,31,32,33,34,35,36,37,38,41]
    $ 1266 "AMR_Done≔ False "
    global AMR_Done=  False
    $ 1267 "AMR_PosActual≔T2O_Current_Pos"
    global AMR_PosActual=modbus_get_signal_status("T2O_Current_Pos")
    $ 1268 "AMR_Attemps≔T2O_Nav_Attemps"
    global AMR_Attemps=modbus_get_signal_status("T2O_Nav_Attemps")
    $ 1269 "AMR_Battery≔MiR_Battery_Lvl"
    global AMR_Battery=modbus_get_signal_status("MiR_Battery_Lvl")
    $ 1270 "AMR_Charging≔(T2O_Charging≟1)"
    global AMR_Charging=(modbus_get_signal_status("T2O_Charging") == 1)
    $ 1271 "AMR_Position≔struct(position_identifier=T2O_Current_Pos, x1=MiR_Position_X1, x2=MiR_Position_X2, y1=MiR_Position_Y1, y2=MiR_Position_Y2, theta1=MiR_Theta_1, theta2=MiR_Theta_2) "
    global AMR_Position=struct(position_identifier=modbus_get_signal_status("T2O_Current_Pos"), x1=modbus_get_signal_status("MiR_Position_X1"), x2=modbus_get_signal_status("MiR_Position_X2"), y1=modbus_get_signal_status("MiR_Position_Y1"), y2=modbus_get_signal_status("MiR_Position_Y2"), theta1=modbus_get_signal_status("MiR_Theta_1"), theta2=modbus_get_signal_status("MiR_Theta_2"))
    $ 1272 "If MiR_Mode≠7"
    if (modbus_get_signal_status("MiR_Mode") != 7):
      $ 1273 "Error"
      $ 1274 "set_error(ERROR_AMR_WRONG_MODE)"
      set_error(ERROR_AMR_WRONG_MODE)
      $ 1275 "AMR_Done≔ True "
      global AMR_Done=  True
    end
    $ 1276 "'=========='"
    # '=========='
    $ 1277 "Switch STATE"
    switch_1 = STATE
    $ 1278 "Case 1"
    if (1 == switch_1):
      $ 1279 "stopping"
      $ 1280 "If T2O_Done≟1 and O2T_Acknowledge≟0"
      if (modbus_get_signal_status("T2O_Done") == 1  and  modbus_get_signal_status("O2T_Acknowledge") == 0):
        $ 1281 "Set O2T_Acknowledge=1"
        modbus_set_output_register("O2T_Acknowledge", 1)
      end
      $ 1282 "Set MiR_CMD_Stop=On"
      modbus_set_output_signal("MiR_CMD_Stop", True)
      $ 1283 "AMR_Position.position_identifier = 0"
      AMR_Position.position_identifier = 0
      $ 1284 "AMR_Done≔ True "
      global AMR_Done=  True
    elif (2 == switch_1):
      $ 1285 "Case 2"
      $ 1286 "stopped"
      $ 1287 "If MiR_State≠3 and MiR_State≠5"
      if (modbus_get_signal_status("MiR_State") != 3  and  modbus_get_signal_status("MiR_State") != 5):
        $ 1288 "Set MiR_CMD_Stop=Off"
        modbus_set_output_signal("MiR_CMD_Stop", False)
      end
    elif (3 == switch_1):
      $ 1289 "Case 3"
      $ 1290 "resetting"
      $ 1291 "Set O2T_Mis_Main=Off"
      modbus_set_output_signal("O2T_Mis_Main", False)
      $ 1292 "Set O2T_Mis_Charge=Off"
      modbus_set_output_signal("O2T_Mis_Charge", False)
      $ 1293 "If MiR_Mis_Queue>0"
      if (modbus_get_signal_status("MiR_Mis_Queue")>0):
        $ 1294 "Set MiR_CMD_Clear_Q=On"
        modbus_set_output_signal("MiR_CMD_Clear_Q", True)
        $ 1295 "Wait MiR_Mis_Queue≟0"
        while (not(modbus_get_signal_status("MiR_Mis_Queue") == 0)):
          sync()
        end
        $ 1296 "Set MiR_CMD_Clear_Q=Off"
        modbus_set_output_signal("MiR_CMD_Clear_Q", False)
      end
      $ 1297 "If MiR_Error_ID≠0"
      if (modbus_get_signal_status("MiR_Error_ID") != 0):
        $ 1298 "Set MiR_CMD_Clear_E=On"
        modbus_set_output_signal("MiR_CMD_Clear_E", True)
        $ 1299 "Wait MiR_Error_ID≟0"
        while (not(modbus_get_signal_status("MiR_Error_ID") == 0)):
          sync()
        end
        $ 1300 "Set MiR_CMD_Clear_E=Off"
        modbus_set_output_signal("MiR_CMD_Clear_E", False)
      end
      $ 1301 "Set O2T_Action=0"
      modbus_set_output_register("O2T_Action", 0)
      $ 1302 "Set O2T_Acknowledge=0"
      modbus_set_output_register("O2T_Acknowledge", 0)
      $ 1303 "Set O2T_Target_Pos=0"
      modbus_set_output_register("O2T_Target_Pos", 0)
      $ 1304 "Set O2T_Footprint=0"
      modbus_set_output_register("O2T_Footprint", 0)
      $ 1305 "Set O2T_ProtectOff=0"
      modbus_set_output_register("O2T_ProtectOff", 0)
      $ 1306 "Set O2T_Dock=0"
      modbus_set_output_register("O2T_Dock", 0)
      $ 1307 "AMR_Attemps≔0"
      global AMR_Attemps=0
      $ 1308 "AMR_PosTarget≔0"
      global AMR_PosTarget=0
      $ 1309 "AMR_Step≔0"
      global AMR_Step=0
      $ 1310 "AMR_AtTarget≔ False "
      global AMR_AtTarget=  False
      $ 1311 "If MiR_State≟4 or MiR_State≟3 or MiR_State≟10"
      if (modbus_get_signal_status("MiR_State") == 4  or  modbus_get_signal_status("MiR_State") == 3  or  modbus_get_signal_status("MiR_State") == 10):
        $ 1312 "AMR_Done≔ True "
        global AMR_Done=  True
      end
    elif (5 == switch_1):
      $ 1313 "Case 5"
      $ 1314 "starting"
      $ 1315 "If MiR_State≟4"
      if (modbus_get_signal_status("MiR_State") == 4):
        $ 1316 "Set MiR_CMD_Start=On"
        modbus_set_output_signal("MiR_CMD_Start", True)
        $ 1317 "Wait MiR_State≠4"
        while (not(modbus_get_signal_status("MiR_State") != 4)):
          sync()
        end
        $ 1318 "Set MiR_CMD_Start=Off"
        modbus_set_output_signal("MiR_CMD_Start", False)
        $ 1319 "AMR_Done≔ True "
        global AMR_Done=  True
      else:
        $ 1320 "ElseIf MiR_State≟10"
        if (modbus_get_signal_status("MiR_State") == 10):
          $ 1321 "'MiR in protective stop. Wait'"
          # 'MiR in protective stop. Wait'
          $ 1322 "AMR_Done≔ True "
          global AMR_Done=  True
        else:
          $ 1323 "ElseIf MiR_State≟3"
          if (modbus_get_signal_status("MiR_State") == 3):
            $ 1324 "AMR_Done≔ True "
            global AMR_Done=  True
          end
        end
      end
    elif (6 == switch_1):
      $ 1325 "Case 6"
      $ 1326 "execute"
      $ 1327 "AMR_AtTarget≔(AMR_PosActual≟AMR_PosTarget)"
      global AMR_AtTarget=(AMR_PosActual == AMR_PosTarget)
      $ 1328 "Switch AMR_Step"
      switch_2 = AMR_Step
      $ 1329 "Case 0"
      if (0 == switch_2):
        $ 1330 "If  not AMR_AtTarget"
        if (  not  AMR_AtTarget):
          $ 1331 "AMR_Step≔1"
          global AMR_Step=1
        else:
          $ 1332 "Else" "noBreak"
          $ 1333 "AMR_Done≔ True "
          global AMR_Done=  True
        end
      elif (1 == switch_2):
        $ 1334 "Case 1"
        $ 1335 "general Settings"
        $ 1336 "Set O2T_Acknowledge=0"
        modbus_set_output_register("O2T_Acknowledge", 0)
        $ 1337 "check for error"
        $ 1338 "If OBJ_Picked and MiR_State≟10"
        if (OBJ_Picked  and  modbus_get_signal_status("MiR_State") == 10):
          $ 1339 "Error"
          $ 1340 "set_error(ERROR_ROBOT_ARM_NOT_IN_HOME_POSE)"
          set_error(ERROR_ROBOT_ARM_NOT_IN_HOME_POSE)
          $ 1341 "Action≔0"
          global Action=0
        else:
          $ 1342 "ElseIf  not found_in_list(AMR_PosTarget, AMR_TargetList)"
          if (  not  found_in_list(AMR_PosTarget, AMR_TargetList)):
            $ 1343 "Error"
            $ 1344 "set_error(ERROR_UNKNOWN_POSE)"
            set_error(ERROR_UNKNOWN_POSE)
            $ 1345 "Action≔0"
            global Action=0
          end
        end
        $ 1346 "If MiR_State≟3"
        if (modbus_get_signal_status("MiR_State") == 3):
          $ 1347 "Set MiR_CMD_Start=Off"
          modbus_set_output_signal("MiR_CMD_Start", False)
          $ 1348 "Switch Action"
          switch_3 = Action
          $ 1349 "Case 51"
          if (51 == switch_3):
            $ 1350 "Charge"
            $ 1351 "'trigger the charging mission'"
            # 'trigger the charging mission'
            $ 1352 "'target pos is predefined'"
            # 'target pos is predefined'
            $ 1353 "Set O2T_Footprint=0"
            modbus_set_output_register("O2T_Footprint", 0)
            $ 1354 "Set O2T_Action=1"
            modbus_set_output_register("O2T_Action", 1)
            $ 1355 "If MiR_Mis_Queue≟0"
            if (modbus_get_signal_status("MiR_Mis_Queue") == 0):
              $ 1356 "Set O2T_Mis_Charge=On"
              modbus_set_output_signal("O2T_Mis_Charge", True)
              $ 1357 "Wait MiR_Mis_Queue≥1"
              while (not(modbus_get_signal_status("MiR_Mis_Queue") >= 1)):
                sync()
              end
              $ 1358 "Set O2T_Mis_Charge=Off"
              modbus_set_output_signal("O2T_Mis_Charge", False)
            end
          elif (52 == switch_3):
            $ 1359 "Case 52"
            $ 1360 "Navigate"
            $ 1361 "'trigger the standard missoin'"
            # 'trigger the standard missoin'
            $ 1362 "Set O2T_Footprint=AMR_FootprintID"
            modbus_set_output_register("O2T_Footprint", AMR_FootprintID)
            $ 1363 "Set O2T_Target_Pos=AMR_PosTarget"
            modbus_set_output_register("O2T_Target_Pos", AMR_PosTarget)
            $ 1364 "Set O2T_Action=2"
            modbus_set_output_register("O2T_Action", 2)
            $ 1365 "If MiR_Mis_Queue≟0"
            if (modbus_get_signal_status("MiR_Mis_Queue") == 0):
              $ 1366 "Set O2T_Mis_Main=On"
              modbus_set_output_signal("O2T_Mis_Main", True)
              $ 1367 "Wait MiR_Mis_Queue≥1"
              while (not(modbus_get_signal_status("MiR_Mis_Queue") >= 1)):
                sync()
              end
              $ 1368 "Set O2T_Mis_Main=Off"
              modbus_set_output_signal("O2T_Mis_Main", False)
            end
          end
        else:
          $ 1369 "ElseIf MiR_State≟4"
          if (modbus_get_signal_status("MiR_State") == 4):
            $ 1370 "Set MiR_CMD_Start=On"
            modbus_set_output_signal("MiR_CMD_Start", True)
          else:
            $ 1371 "ElseIf MiR_State≟5"
            if (modbus_get_signal_status("MiR_State") == 5):
              $ 1372 "AMR_Step≔2"
              global AMR_Step=2
            else:
              $ 1373 "ElseIf MiR_State≟10"
              if (modbus_get_signal_status("MiR_State") == 10):
                $ 1374 "'AMR still in safeguard stop'"
                # 'AMR still in safeguard stop'
              end
            end
          end
        end
      elif (2 == switch_2):
        $ 1375 "Case 2"
        $ 1376 "acknowledge handshake"
        $ 1377 "If T2O_Done≟1 and O2T_Acknowledge≟0"
        if (modbus_get_signal_status("T2O_Done") == 1  and  modbus_get_signal_status("O2T_Acknowledge") == 0):
          $ 1378 "Set O2T_Acknowledge=1"
          modbus_set_output_register("O2T_Acknowledge", 1)
        else:
          $ 1379 "ElseIf T2O_Done≟0 and O2T_Acknowledge≟1"
          if (modbus_get_signal_status("T2O_Done") == 0  and  modbus_get_signal_status("O2T_Acknowledge") == 1):
            $ 1380 "Set O2T_Acknowledge=0"
            modbus_set_output_register("O2T_Acknowledge", 0)
            $ 1381 "AMR_AtTarget≔(AMR_PosActual≟AMR_PosTarget)"
            global AMR_AtTarget=(AMR_PosActual == AMR_PosTarget)
            $ 1382 "AMR_Done≔ True "
            global AMR_Done=  True
          end
        end
      end
      $ 1383 "translate errors"
      $ 1384 "If AMR_Done"
      if (AMR_Done):
        $ 1385 "Switch T2O_Error_ID"
        switch_2 = modbus_get_signal_status("T2O_Error_ID")
        $ 1386 "Case 2003"
        if (2003 == switch_2):
          $ 1387 "error"
          $ 1388 "set_error(ERROR_NOT_DOCKED)"
          set_error(ERROR_NOT_DOCKED)
        elif (2007 == switch_2):
          $ 1389 "Case 2007"
          $ 1390 "error"
          $ 1391 "set_error(ERROR_NOT_REACHABLE_TARGET)"
          set_error(ERROR_NOT_REACHABLE_TARGET)
        elif (2008 == switch_2):
          $ 1392 "Case 2008"
          $ 1393 "error"
          $ 1394 "set_error(ERROR_CHARGING_NOT_STARTED)"
          set_error(ERROR_CHARGING_NOT_STARTED)
        end
      end
    elif (7 == switch_1):
      $ 1395 "Case 7"
      $ 1396 "completing"
      $ 1397 "If MiR_Mis_Queue>0"
      if (modbus_get_signal_status("MiR_Mis_Queue")>0):
        $ 1398 "Set MiR_CMD_Abort=On"
        modbus_set_output_signal("MiR_CMD_Abort", True)
        $ 1399 "Wait MiR_Mis_Queue≟0"
        while (not(modbus_get_signal_status("MiR_Mis_Queue") == 0)):
          sync()
        end
        $ 1400 "Set MiR_CMD_Abort=Off"
        modbus_set_output_signal("MiR_CMD_Abort", False)
      end
      $ 1401 "If MiR_State≟3 or MiR_State≟10"
      if (modbus_get_signal_status("MiR_State") == 3  or  modbus_get_signal_status("MiR_State") == 10):
        $ 1402 "AMR_Done≔ True "
        global AMR_Done=  True
      end
    elif (9 == switch_1):
      $ 1403 "Case 9"
      $ 1404 "holding"
      $ 1405 "Set MiR_CMD_Abort=On"
      modbus_set_output_signal("MiR_CMD_Abort", True)
      $ 1406 "If MiR_State≟3 or MiR_State≟10"
      if (modbus_get_signal_status("MiR_State") == 3  or  modbus_get_signal_status("MiR_State") == 10):
        $ 1407 "Set MiR_CMD_Abort=Off"
        modbus_set_output_signal("MiR_CMD_Abort", False)
        $ 1408 "AMR_Done≔ True "
        global AMR_Done=  True
      end
    elif (11 == switch_1):
      $ 1409 "Case 11"
      $ 1410 "unholding"
      $ 1411 "Set MiR_CMD_Start=On"
      modbus_set_output_signal("MiR_CMD_Start", True)
      $ 1412 "If MiR_State≠4"
      if (modbus_get_signal_status("MiR_State") != 4):
        $ 1413 "Set MiR_CMD_Start=Off"
        modbus_set_output_signal("MiR_CMD_Start", False)
        $ 1414 "AMR_Step≔0"
        global AMR_Step=0
        $ 1415 "AMR_Done≔ True "
        global AMR_Done=  True
      end
    elif (12 == switch_1):
      $ 1416 "Case 12"
      $ 1417 "suspending"
      $ 1418 "'none'"
      # 'none'
    elif (14 == switch_1):
      $ 1419 "Case 14"
      $ 1420 "unsuspending"
      $ 1421 "'none'"
      # 'none'
    elif (15 == switch_1):
      $ 1422 "Case 15"
      $ 1423 "aborting"
      $ 1424 "Set MiR_CMD_Abort=On"
      modbus_set_output_signal("MiR_CMD_Abort", True)
      $ 1425 "Wait MiR_State≟3"
      while (not(modbus_get_signal_status("MiR_State") == 3)):
        sync()
      end
      $ 1426 "Set MiR_CMD_Abort=Off"
      modbus_set_output_signal("MiR_CMD_Abort", False)
    elif (17 == switch_1):
      $ 1427 "Case 17"
      $ 1428 "clearing"
      $ 1429 "If MiR_Error_ID≠0"
      if (modbus_get_signal_status("MiR_Error_ID") != 0):
        $ 1430 "Set MiR_CMD_Clear_E=On"
        modbus_set_output_signal("MiR_CMD_Clear_E", True)
        $ 1431 "Wait MiR_Error_ID≟0"
        while (not(modbus_get_signal_status("MiR_Error_ID") == 0)):
          sync()
        end
        $ 1432 "Set MiR_CMD_Clear_E=Off"
        modbus_set_output_signal("MiR_CMD_Clear_E", False)
      end
      $ 1433 "If MiR_Error_ID≟0"
      if (modbus_get_signal_status("MiR_Error_ID") == 0):
        $ 1434 "AMR_Done≔ True "
        global AMR_Done=  True
      end
    end
    $ 1435 "'=========='"
    # '=========='
    $ 1436 "PostSettings"
    $ 1437 "AMR_Position≔struct(position_identifier=T2O_Current_Pos, x1=MiR_Position_X1, x2=MiR_Position_X2, y1=MiR_Position_Y1, y2=MiR_Position_Y2, theta1=MiR_Theta_1, theta2=MiR_Theta_2) "
    global AMR_Position=struct(position_identifier=modbus_get_signal_status("T2O_Current_Pos"), x1=modbus_get_signal_status("MiR_Position_X1"), x2=modbus_get_signal_status("MiR_Position_X2"), y1=modbus_get_signal_status("MiR_Position_Y1"), y2=modbus_get_signal_status("MiR_Position_Y2"), theta1=modbus_get_signal_status("MiR_Theta_1"), theta2=modbus_get_signal_status("MiR_Theta_2"))
  end
  def Sub_Action_V4():
    $ 1438 "Sub_Action_V4" "noBreak"
    $ 1439 "PreSettings"
    $ 1440 "init poses"
    $ 1441 "PSE_A≔p[0,0,0,0,0,0]"
    global PSE_A=p[0,0,0,0,0,0]
    $ 1442 "PSE_A_H≔p[0,0,0,0,0,0]"
    global PSE_A_H=p[0,0,0,0,0,0]
    $ 1443 "PSE_T≔p[0,0,0,0,0,0]"
    global PSE_T=p[0,0,0,0,0,0]
    $ 1444 "PSE_T_H≔p[0,0,0,0,0,0]"
    global PSE_T_H=p[0,0,0,0,0,0]
    $ 1445 "PSE_G≔p[0,0,0,0,0,0]"
    global PSE_G=p[0,0,0,0,0,0]
    $ 1446 "PSE_G_H≔p[0,0,0,0,0,0]"
    global PSE_G_H=p[0,0,0,0,0,0]
    $ 1447 "PSE_R≔p[0,0,0,0,0,0]"
    global PSE_R=p[0,0,0,0,0,0]
    $ 1448 "PSE_R_H≔p[0,0,0,0,0,0]"
    global PSE_R_H=p[0,0,0,0,0,0]
    $ 1449 "JNT_Q≔[0,0,0,0,0,0]"
    global JNT_Q=[0,0,0,0,0,0]
    $ 1450 "JNT_S≔[0,0,0,0,0,0]"
    global JNT_S=[0,0,0,0,0,0]
    $ 1451 "Gripping parameters"
    $ 1452 "OBJ = find_object_by_type(OBJs, OBJ_Type)"
    OBJ = find_object_by_type(OBJs, OBJ_Type)
    $ 1453 "GRP_Open_Pos≔OBJ.dimension.diameter * 1000 + 6"
    global GRP_Open_Pos=OBJ.dimension.diameter * 1000 + 6
    $ 1454 "GRP_Offset≔OBJ.gripper_offset"
    global GRP_Offset=OBJ.gripper_offset
    $ 1455 "rq_set_force_norm(50)"
     rq_set_force_norm (50)
    $ 1456 "rq_set_speed_norm(50)"
     rq_set_speed_norm (50)
    $ 1457 "Switch ITM_ID"
    switch_1 = ITM_ID
    $ 1458 "Case 1"
    if (1 == switch_1):
      $ 1459 "uML"
      $ 1460 "JIG2 = find_object_by_type(JIGs, JIG)"
      JIG2 = find_object_by_type(JIGs, JIG)
      $ 1461 "JIG_Offset≔JIG2.jig_offset"
      global JIG_Offset=JIG2.jig_offset
      $ 1462 "Switch JIG"
      switch_2 = JIG
      $ 1463 "Case 1"
      if (1 == switch_2):
        $ 1464 "3FG"
        $ 1465 "define poses"
        $ 1466 "FRM_Reference≔ULM_3FG"
        global FRM_Reference=ULM_3FG
        $ 1467 "JNT_Q≔JNT_HOME"
        global JNT_Q=JNT_HOME
        $ 1468 "PSE_T≔pose_trans(GRP_Offset, JIG_Offset)"
        global PSE_T= pose_trans (GRP_Offset, JIG_Offset)
        $ 1469 "PSE_A≔pose_trans(PSE_T, p[0,0,0.100,0,0,0])"
        global PSE_A= pose_trans (PSE_T, p[0,0,0.100,0,0,0])
        $ 1470 "PSE_R≔pose_add(PSE_T, p[0,0,0.100,0,0,0])"
        global PSE_R= pose_add (PSE_T, p[0,0,0.100,0,0,0])
      elif (2 == switch_2):
        $ 1471 "Case 2"
        $ 1472 "Input"
        $ 1473 "'CHANGE THE REFERENCE TO THE FRAME TO MOVE IN'"
        # 'CHANGE THE REFERENCE TO THE FRAME TO MOVE IN'
        $ 1474 "define poses"
        $ 1475 "FRM_Reference≔ULM_Input"
        global FRM_Reference=ULM_Input
        $ 1476 "PSE_T≔pose_trans(pose_trans(get_pattern_pos_rectangle(OBJ_Nbr, 'X', [10,5], patternsize=[0.181,0.081]), GRP_Offset), JIG_Offset)"
        global PSE_T= pose_trans ( pose_trans (get_pattern_pos_rectangle(OBJ_Nbr, "X", [10,5], patternsize=[0.181,0.081]), GRP_Offset), JIG_Offset)
        $ 1477 "If Action≟1"
        if (Action == 1):
          $ 1478 "PSE_R≔pose_add(PSE_T, p[0,0,0.200,0,0,0])"
          global PSE_R= pose_add (PSE_T, p[0,0,0.200,0,0,0])
          $ 1479 "PSE_A≔pose_add(PSE_T, p[0,0,0.100,0,0,0])"
          global PSE_A= pose_add (PSE_T, p[0,0,0.100,0,0,0])
        else:
          $ 1480 "ElseIf Action≟2"
          if (Action == 2):
            $ 1481 "PSE_R≔pose_add(PSE_T, p[0,0,0.100,0,0,0])"
            global PSE_R= pose_add (PSE_T, p[0,0,0.100,0,0,0])
            $ 1482 "PSE_A≔pose_add(PSE_T, p[0,0,0.200,0,0,0])"
            global PSE_A= pose_add (PSE_T, p[0,0,0.200,0,0,0])
          end
        end
      elif (3 == switch_2):
        $ 1483 "Case 3"
        $ 1484 "Output"
        $ 1485 "'CHANGE THE REFERENCE TO THE FRAME TO MOVE IN'"
        # 'CHANGE THE REFERENCE TO THE FRAME TO MOVE IN'
        $ 1486 "define poses"
        $ 1487 "FRM_Reference≔ULM_Output"
        global FRM_Reference=ULM_Output
        $ 1488 "PSE_T≔pose_trans(pose_trans(get_pattern_pos_rectangle(OBJ_Nbr, 'X', [10,5], patternsize=[0.181,0.081]), GRP_Offset), JIG_Offset)"
        global PSE_T= pose_trans ( pose_trans (get_pattern_pos_rectangle(OBJ_Nbr, "X", [10,5], patternsize=[0.181,0.081]), GRP_Offset), JIG_Offset)
        $ 1490 "If Action≟1"
        if (Action == 1):
          $ 1491 "PSE_R≔pose_add(PSE_T, p[0,0,0.200,0,0,0])"
          global PSE_R= pose_add (PSE_T, p[0,0,0.200,0,0,0])
          $ 1492 "PSE_A≔pose_add(PSE_T, p[0,0,0.100,0,0,0])"
          global PSE_A= pose_add (PSE_T, p[0,0,0.100,0,0,0])
        else:
          $ 1493 "ElseIf Action≟2"
          if (Action == 2):
            $ 1494 "PSE_R≔pose_add(PSE_T, p[0,0,0.100,0,0,0])"
            global PSE_R= pose_add (PSE_T, p[0,0,0.100,0,0,0])
            $ 1495 "PSE_A≔pose_add(PSE_T, p[0,0,0.200,0,0,0])"
            global PSE_A= pose_add (PSE_T, p[0,0,0.200,0,0,0])
          end
        end
      elif (4 == switch_2):
        $ 1496 "Case 4"
        $ 1497 "jig centrifuge racks"
        $ 1498 "define poses"
        $ 1499 "FRM_Reference≔ULM_Cent_Racks"
        global FRM_Reference=ULM_Cent_Racks
        $ 1500 "PSE_T≔get_pattern_pos_rectangle(JIG_Slot, 'X', [4,1], patternsize=[0.291,0])"
        global PSE_T=get_pattern_pos_rectangle(JIG_Slot, "X", [4,1], patternsize=[0.291,0])
        $ 1501 "If OBJ_Nbr≠0"
        if (OBJ_Nbr != 0):
          $ 1502 "PSE_T≔pose_trans(pose_trans(PSE_T, get_pattern_pos_rectangle(OBJ_Nbr, 'X', [3,3], patternsize=[0.060,0.060])),p[-0.030, -0.030,0,0,0,3.927])"
          global PSE_T= pose_trans ( pose_trans (PSE_T, get_pattern_pos_rectangle(OBJ_Nbr, "X", [3,3], patternsize=[0.060,0.060])),p[-0.030, -0.030,0,0,0,3.927])
        end
        $ 1503 "PSE_T≔pose_trans(PSE_T, GRP_Offset)"
        global PSE_T= pose_trans (PSE_T, GRP_Offset)
        $ 1504 "If Action≟1"
        if (Action == 1):
          $ 1505 "PSE_R≔pose_add(PSE_T, p[0,0,0.200,0,0,0])"
          global PSE_R= pose_add (PSE_T, p[0,0,0.200,0,0,0])
          $ 1506 "PSE_A≔pose_add(PSE_T, p[0,0,0.100,0,0,0])"
          global PSE_A= pose_add (PSE_T, p[0,0,0.100,0,0,0])
        else:
          $ 1507 "ElseIf Action≟2"
          if (Action == 2):
            $ 1508 "PSE_R≔pose_add(PSE_T, p[0,0,0.100,0,0,0])"
            global PSE_R= pose_add (PSE_T, p[0,0,0.100,0,0,0])
            $ 1509 "PSE_A≔pose_add(PSE_T, p[0,0,0.200,0,0,0])"
            global PSE_A= pose_add (PSE_T, p[0,0,0.200,0,0,0])
          end
        end
      elif (6 == switch_2):
        $ 1510 "Case 6"
        $ 1511 "Caps bin"
        $ 1512 "define poses"
        $ 1513 "'Drop cap'"
        # 'Drop cap'
        $ 1514 "FRM_Reference=ULM_Cap_Bin"
        FRM_Reference=ULM_Cap_Bin
        $ 1515 "PSE_T≔pose_RPY2RotVec(p[0,0,0,0,0,0])"
        global PSE_T=pose_RPY2RotVec(p[0,0,0,0,0,0])
        $ 1516 "PSE_T_H≔pose_add(PSE_T, p[0,0,-0.011,0,0,0])"
        global PSE_T_H= pose_add (PSE_T, p[0,0,-0.011,0,0,0])
        $ 1517 "PSE_A≔pose_trans(PSE_T, p[0,0,0.1,0,0,0])"
        global PSE_A= pose_trans (PSE_T, p[0,0,0.1,0,0,0])
        $ 1518 "PSE_R_H≔pose_add(PSE_T, p[0,0,0.100,0,0,0])"
        global PSE_R_H= pose_add (PSE_T, p[0,0,0.100,0,0,0])
        $ 1519 "PSE_R≔pose_add(PSE_T, p[0,0,0.100,0,0,0])"
        global PSE_R= pose_add (PSE_T, p[0,0,0.100,0,0,0])
      elif (7 == switch_2):
        $ 1520 "Case 7"
        $ 1521 "Sarstedt"
        $ 1522 "'CHANGE THE REFERENCE TO THE FRAME TO MOVE IN'"
        # 'CHANGE THE REFERENCE TO THE FRAME TO MOVE IN'
        $ 1528 "If TASK.ID≟10"
        if (TASK.ID == 10):
          $ 1529 "Frame & Position Params"
          $ 1531 "FRM_Reference = CAM_LM_SSRack"
          FRM_Reference = CAM_LM_SSRack
          $ 1536 "PSE_T≔uLM_SS_PickPlc"
          global PSE_T=uLM_SS_PickPlc
          $ 1537 "PSE_A≔pose_trans(PSE_T, p[0,0,0.1,0,0,0])"
          global PSE_A= pose_trans (PSE_T, p[0,0,0.1,0,0,0])
          $ 1538 "PSE_R≔pose_add(PSE_T, p[0,0,0.1,0,0,0])"
          global PSE_R= pose_add (PSE_T, p[0,0,0.1,0,0,0])
        else:
          $ 1539 "ElseIf TASK.ID≟11"
          if (TASK.ID == 11):
            $ 1540 "FRM_Reference = ULM_SS_Jig"
            FRM_Reference = ULM_SS_Jig
            $ 1541 "PSE_T≔pose_RPY2RotVec(p[0,0,0,0,0,0])"
            global PSE_T=pose_RPY2RotVec(p[0,0,0,0,0,0])
            $ 1542 "PSE_T≔pose_trans(PSE_T, GRP_Offset)"
            global PSE_T=pose_trans(PSE_T, GRP_Offset)
            $ 1543 "PSE_A≔pose_trans(PSE_T, p[0,0,0.1,0,0,0])"
            global PSE_A= pose_trans (PSE_T, p[0,0,0.1,0,0,0])
            $ 1544 "PSE_R≔pose_add(PSE_T, p[0,0,0.2,0,0,0])"
            global PSE_R= pose_add (PSE_T, p[0,0,0.2,0,0,0])
          end
        end
      elif (8 == switch_2):
        $ 1545 "Case 8"
        $ 1546 "NoK"
        $ 1547 "define poses"
        $ 1548 "'NoK'"
        # 'NoK'
        $ 1549 "FRM_Reference=ULM_NoK"
        FRM_Reference=ULM_NoK
        $ 1550 "PSE_T≔pose_RPY2RotVec(p[0,0,0,0,0,0])"
        global PSE_T=pose_RPY2RotVec(p[0,0,0,0,0,0])
        $ 1551 "PSE_A≔pose_trans(PSE_T, p[0,0,0.1,0,0,0])"
        global PSE_A= pose_trans (PSE_T, p[0,0,0.1,0,0,0])
        $ 1552 "PSE_R≔pose_add(PSE_T, p[0,0,0.100,0,0,0])"
        global PSE_R= pose_add (PSE_T, p[0,0,0.100,0,0,0])
      elif (9 == switch_2):
        $ 1553 "Case 9"
        $ 1554 "Pick_bott_jig"
        $ 1555 "define poses"
        $ 1556 "'NoK'"
        # 'NoK'
        $ 1557 "FRM_Reference=ULM_bottle_pick_const"
        FRM_Reference=p[0.08175869478771049,-0.47602162643540935,0.09,0.00141829700319658,-0.0027789445191063835,0.07763675748118615]
        $ 1558 "PSE_T≔pose_RPY2RotVec(p[0,0,0,0,0,0])"
        global PSE_T=pose_RPY2RotVec(p[0,0,0,0,0,0])
        $ 1559 "PSE_A≔pose_trans(PSE_T, p[0,0,0.1,0,0,0])"
        global PSE_A= pose_trans (PSE_T, p[0,0,0.1,0,0,0])
        $ 1560 "PSE_R≔pose_add(PSE_T, p[0,0,0.100,0,0,0])"
        global PSE_R= pose_add (PSE_T, p[0,0,0.100,0,0,0])
      elif (10 == switch_2):
        $ 1561 "Case 10"
        $ 1562 "Place_bott_jig"
        $ 1563 "define poses"
        $ 1564 "'NoK'"
        # 'NoK'
        $ 1565 "FRM_Reference=ULM_bottle_plac_const"
        FRM_Reference=p[-0.09502738395762109,-0.5154087721098056,0.095,0.0014590126708889871,-0.0028280855286173575,0.07763149296298452]
        $ 1566 "PSE_T≔pose_RPY2RotVec(p[0,0,0,0,0,0])"
        global PSE_T=pose_RPY2RotVec(p[0,0,0,0,0,0])
        $ 1567 "PSE_A≔pose_trans(PSE_T, p[0,0,0.1,0,0,0])"
        global PSE_A= pose_trans (PSE_T, p[0,0,0.1,0,0,0])
        $ 1568 "PSE_R≔pose_add(PSE_T, p[0,0,0.100,0,0,0])"
        global PSE_R= pose_add (PSE_T, p[0,0,0.100,0,0,0])
      elif (11 == switch_2):
        $ 1569 "Case 11"
        $ 1570 "Place_bott_jig"
        $ 1571 "define poses"
        $ 1572 "'NoK'"
        # 'NoK'
        $ 1573 "FRM_Reference=shake"
        FRM_Reference=shake
        $ 1574 "PSE_T≔pose_RPY2RotVec(p[0,0,0,0,0,0])"
        global PSE_T=pose_RPY2RotVec(p[0,0,0,0,0,0])
        $ 1575 "PSE_A≔pose_trans(PSE_T, p[0,0,0,0,0,0])"
        global PSE_A= pose_trans (PSE_T, p[0,0,0,0,0,0])
        $ 1576 "PSE_R≔pose_add(PSE_T, p[0,0,0,0,0,0])"
        global PSE_R= pose_add (PSE_T, p[0,0,0,0,0,0])
      elif (12 == switch_2):
        $ 1577 "Case 12"
        $ 1578 "Pick_Vial_jig"
        $ 1579 "define poses"
        $ 1580 "'NoK'"
        # 'NoK'
        $ 1581 "FRM_Reference=shake"
        FRM_Reference=shake
        $ 1582 "PSE_T≔pose_RPY2RotVec(p[0,0,0,0,0,0])"
        global PSE_T=pose_RPY2RotVec(p[0,0,0,0,0,0])
        $ 1583 "PSE_A≔pose_trans(PSE_T, p[0,0,0,0,0,0])"
        global PSE_A= pose_trans (PSE_T, p[0,0,0,0,0,0])
        $ 1584 "PSE_R≔pose_add(PSE_T, p[0,0,0,0,0,0])"
        global PSE_R= pose_add (PSE_T, p[0,0,0,0,0,0])
      end
    elif (2 == switch_1):
      $ 1585 "Case 2"
      $ 1586 "Centrifuge"
      $ 1587 "'CHANGE THE REFERENCE TO THE FRAME TO MOVE IN'"
      # 'CHANGE THE REFERENCE TO THE FRAME TO MOVE IN'
      $ 1588 "define poses"
      $ 1589 "FRM_Reference≔FRM_Centrifuge"
      global FRM_Reference=FRM_Centrifuge
      $ 1590 "PSE_T≔GRP_Offset"
      global PSE_T=GRP_Offset
      $ 1591 "If Action≟8"
      if (Action == 8):
        $ 1592 "PSE_R≔pose_add(PSE_T, p[0,0,0.250,0,0,0])"
        global PSE_R= pose_add (PSE_T, p[0,0,0.250,0,0,0])
        $ 1593 "PSE_A≔pose_add(PSE_T, p[0,0,0.150,0,0,0])"
        global PSE_A= pose_add (PSE_T, p[0,0,0.150,0,0,0])
      else:
        $ 1594 "ElseIf Action≟7"
        if (Action == 7):
          $ 1595 "PSE_R≔pose_add(PSE_T, p[0,0,0.150,0,0,0])"
          global PSE_R= pose_add (PSE_T, p[0,0,0.150,0,0,0])
          $ 1596 "PSE_A≔pose_add(PSE_T, p[0,0,0.250,0,0,0])"
          global PSE_A= pose_add (PSE_T, p[0,0,0.250,0,0,0])
        end
      end
    elif (3 == switch_1):
      $ 1597 "Case 3"
      $ 1598 "Output"
      $ 1599 "'CHANGE THE REFERENCE TO THE FRAME TO MOVE IN'"
      # 'CHANGE THE REFERENCE TO THE FRAME TO MOVE IN'
      $ 1600 "define poses"
      $ 1601 "FRM_Reference≔Base_const"
      global FRM_Reference=p[0.0,0.0,0.0,0.0,0.0,0.0]
      $ 1602 "PSE_T≔p[0,0,0,0,0,0]"
      global PSE_T=p[0,0,0,0,0,0]
      $ 1603 "PSE_A≔pose_add(PSE_T, p[0,0,0.150,0,0,0])"
      global PSE_A= pose_add (PSE_T, p[0,0,0.150,0,0,0])
      $ 1604 "PSE_R≔pose_add(PSE_T, p[0,0,0.100,0,0,0])"
      global PSE_R= pose_add (PSE_T, p[0,0,0.100,0,0,0])
    elif (5 == switch_1):
      $ 1605 "Case 5"
      $ 1606 "Sarstedt Pickup Table"
      $ 1607 "'CHANGE THE REFERENCE TO THE FRAME TO MOVE IN'"
      # 'CHANGE THE REFERENCE TO THE FRAME TO MOVE IN'
      $ 1608 "Switch JIG"
      switch_2 = JIG
      $ 1609 "Case 7"
      if (7 == switch_2):
        $ 1622 "Sarstedt"
        $ 1623 "'CHANGE THE REFERENCE TO THE FRAME TO MOVE IN'"
        # 'CHANGE THE REFERENCE TO THE FRAME TO MOVE IN'
        $ 1629 "If TASK.ID≟10"
        if (TASK.ID == 10):
          $ 1630 "Frame & Position Params"
          $ 1631 "FRM_Reference = CAM_LM_SSRack"
          FRM_Reference = CAM_LM_SSRack
          $ 1632 "PSE_T≔uLM_SS_PickPlc"
          global PSE_T=uLM_SS_PickPlc
          $ 1633 "PSE_A≔pose_trans(PSE_T, p[0,0,0.1,0,0,0])"
          global PSE_A= pose_trans (PSE_T, p[0,0,0.1,0,0,0])
          $ 1634 "PSE_R≔pose_add(PSE_T, p[0,0,0.1,0,0,0])"
          global PSE_R= pose_add (PSE_T, p[0,0,0.1,0,0,0])
        end
      end
    elif (13 == switch_1):
      $ 1641 "Case 13"
      $ 1642 "Sarstedt Pickup Table"
      $ 1643 "'CHANGE THE REFERENCE TO THE FRAME TO MOVE IN'"
      # 'CHANGE THE REFERENCE TO THE FRAME TO MOVE IN'
      $ 1644 "Switch JIG"
      switch_2 = JIG
      $ 1645 "Case 7"
      if (7 == switch_2):
        $ 1658 "Bottle"
        $ 1659 "'CHANGE THE REFERENCE TO THE FRAME TO MOVE IN'"
        # 'CHANGE THE REFERENCE TO THE FRAME TO MOVE IN'
        $ 1665 "If TASK.ID≟43"
        if (TASK.ID == 43):
          $ 1666 "Frame & Position Params"
          $ 1667 "FRM_Reference = CAM_LM_Bott"
          FRM_Reference = CAM_LM_Bott
          $ 1668 "PSE_T≔uLM_SS_PickPlc"
          global PSE_T=uLM_SS_PickPlc
          $ 1669 "PSE_A≔pose_trans(PSE_T, p[0,0,0.1,0,0,0])"
          global PSE_A= pose_trans (PSE_T, p[0,0,0.1,0,0,0])
          $ 1670 "PSE_R≔pose_add(PSE_T, p[0,0,0.1,0,0,0])"
          global PSE_R= pose_add (PSE_T, p[0,0,0.1,0,0,0])
        end
      end
    end
    $ 1677 "Additional check"
    $ 1678 "If  not is_reachable(FRM_Reference,[PSE_A,PSE_A_H,PSE_T,PSE_T_H,PSE_R,PSE_R_H])"
    if (  not  is_reachable(FRM_Reference,[PSE_A,PSE_A_H,PSE_T,PSE_T_H,PSE_R,PSE_R_H])):
      $ 1679 "Error"
      $ 1680 "set_error(ERROR_POSE_NOT_REACHABLE)"
      set_error(ERROR_POSE_NOT_REACHABLE)
      $ 1681 "Action≔0"
      global Action=0
    end
    $ 1682 "'=========='"
    # '=========='
    $ 1683 "Switch Action"
    switch_1 = Action
    $ 1684 "Case 1"
    if (1 == switch_1):
      $ 1685 "Pick"
      $ 1686 "Action_Info≔'pick object'"
      global Action_Info="pick object"
      $ 1687 "do_transition(pose_trans(FRM_Reference, PSE_T), keep_rxry=OBJ_Picked)"
      do_transition( pose_trans (FRM_Reference, PSE_T), keep_rxry=OBJ_Picked)
      $ 1688 "EOAT"
      $ 1689 "If  not OBJ_Picked"
      if (  not  OBJ_Picked):
        $ 1690 "rq_move_and_wait_mm(GRP_Open_Pos)"
         rq_move_and_wait_mm (GRP_Open_Pos)
      end
      $ 1691 "If PSE_A_H≠PSE_Z"
      if (PSE_A_H != PSE_Z):
        $ 1692 "If JNT_Q≠JNT_Z"
        if (JNT_Q != JNT_Z):
          $ 1693 "movej(get_inverse_kin(pose_trans(FRM_Reference, PSE_A_H), qnear=JNT_Q), r=0.050)"
          movej(get_inverse_kin( pose_trans (FRM_Reference, PSE_A_H), qnear=JNT_Q), r=0.050)
        else:
          $ 1694 "Else" "noBreak"
          $ 1695 "movej(pose_trans(FRM_Reference, PSE_A_H), r=0.050)"
          movej( pose_trans (FRM_Reference, PSE_A_H), r=0.050)
        end
      end
      $ 1696 "If PSE_A≠PSE_Z"
      if (PSE_A != PSE_Z):
        $ 1697 "If JNT_Q≠JNT_Z"
        if (JNT_Q != JNT_Z):
          $ 1698 "movej(get_inverse_kin(pose_trans(FRM_Reference, PSE_A), qnear=JNT_Q), r=0.020)"
          movej(get_inverse_kin( pose_trans (FRM_Reference, PSE_A), qnear=JNT_Q), r=0.020)
        else:
          $ 1699 "Else" "noBreak"
          $ 1700 "movej(pose_trans(FRM_Reference, PSE_A), r=0.020)"
          movej( pose_trans (FRM_Reference, PSE_A), r=0.020)
        end
      end
      $ 1701 "MoveL"
      $ 1702 "If PSE_T_H≠PSE_Z"
      if (PSE_T_H != PSE_Z):
        $ 1703 "PSE_T_H" "breakAfter"
        movel(pose_trans(FRM_Reference, PSE_T_H), a=0.5, v=0.4, r=0.01)
      end
      $ 1704 "PSE_T" "breakAfter"
      movel(pose_trans(FRM_Reference, PSE_T), a=0.08, v=0.12)
      $ 1705 "EOAT"
      $ 1706 "rq_set_force_norm(50)"
       rq_set_force_norm (50)
      $ 1707 "rq_close_and_wait()"
       rq_close_and_wait ()
      $ 1708 "OBJ_Picked≔rq_is_object_detected()"
      global OBJ_Picked= rq_is_object_detected ()
      $ 1709 "If  not OBJ_Picked"
      if (  not  OBJ_Picked):
        $ 1710 "set_error(ERROR_NO_OBJECT_TO_PICK)"
        set_error(ERROR_NO_OBJECT_TO_PICK)
      end
      $ 1711 "EXTT"
      $ 1712 "Switch JIG"
      switch_2 = JIG
      $ 1713 "Case 1"
      if (1 == switch_2):
        $ 1714 "3FG"
        $ 1715 "If OBJ_Picked"
        if (OBJ_Picked):
          $ 1716 "Set GRP_3F_Open=On"
          set_standard_digital_out(5, True)
        end
      end
      $ 1717 "If PSE_R_H≠PSE_Z"
      if (PSE_R_H != PSE_Z):
        $ 1718 "PSE_R" "breakAfter"
        movel(pose_trans(FRM_Reference, PSE_R), a=0.5, v=0.4, r=0.01)
        $ 1719 "PSE_R_H" "breakAfter"
        movel(pose_trans(FRM_Reference, PSE_R_H), a=0.5, v=0.4)
      else:
        $ 1720 "Else" "noBreak"
        $ 1721 "PSE_R" "breakAfter"
        movel(pose_trans(FRM_Reference, PSE_R), a=0.5, v=0.4)
      end
    elif (2 == switch_1):
      $ 1722 "Case 2"
      $ 1723 "Place"
      $ 1724 "Action_Info≔'place object'"
      global Action_Info="place object"
      $ 1725 "do_transition(pose_trans(FRM_Reference, PSE_T), keep_rxry=OBJ_Picked)"
      do_transition( pose_trans (FRM_Reference, PSE_T), keep_rxry=OBJ_Picked)
      $ 1726 "EXTT"
      $ 1727 "Switch JIG"
      switch_2 = JIG
      $ 1728 "Case 1"
      if (1 == switch_2):
        $ 1729 "3FG"
        $ 1730 "If OBJ_Picked"
        if (OBJ_Picked):
          $ 1731 "Set GRP_3F_Open=On"
          set_standard_digital_out(5, True)
        end
      end
      $ 1732 "If PSE_A_H≠PSE_Z"
      if (PSE_A_H != PSE_Z):
        $ 1733 "If JNT_Q≠JNT_Z"
        if (JNT_Q != JNT_Z):
          $ 1734 "movej(get_inverse_kin(pose_trans(FRM_Reference, PSE_A_H), qnear=JNT_Q), r=0.050)"
          movej(get_inverse_kin( pose_trans (FRM_Reference, PSE_A_H), qnear=JNT_Q), r=0.050)
        else:
          $ 1735 "Else" "noBreak"
          $ 1736 "movej(pose_trans(FRM_Reference, PSE_A_H), r=0.050)"
          movej( pose_trans (FRM_Reference, PSE_A_H), r=0.050)
        end
      end
      $ 1737 "If PSE_A≠PSE_Z"
      if (PSE_A != PSE_Z):
        $ 1738 "If JNT_Q≠JNT_Z"
        if (JNT_Q != JNT_Z):
          $ 1739 "movej(get_inverse_kin(pose_trans(FRM_Reference, PSE_A), qnear=JNT_Q), r=0.020)"
          movej(get_inverse_kin( pose_trans (FRM_Reference, PSE_A), qnear=JNT_Q), r=0.020)
        else:
          $ 1740 "Else" "noBreak"
          $ 1741 "movej(pose_trans(FRM_Reference, PSE_A), r=0.020)"
          movej( pose_trans (FRM_Reference, PSE_A), r=0.020)
        end
      end
      $ 1742 "MoveL"
      $ 1743 "If PSE_T_H≠PSE_Z"
      if (PSE_T_H != PSE_Z):
        $ 1744 "PSE_T_H" "breakAfter"
        movel(pose_trans(FRM_Reference, PSE_T_H), a=0.5, v=0.4, r=0.01)
      end
      $ 1745 "PSE_T" "breakAfter"
      global move_thread_flag_1745=0
      thread move_thread_1745():
        enter_critical
        move_thread_flag_1745 = 1
        movel(pose_trans(FRM_Reference, PSE_T), a=0.05, v=0.09)
        move_thread_flag_1745 = 2
        exit_critical
      end
      move_thread_flag_1745 = 0
      move_thread_han_1745 = run move_thread_1745()
      while (True):
        local targetTcpDirection=get_target_tcp_speed()
        local stepsToRetract=tool_contact(direction=targetTcpDirection)
        if (stepsToRetract > 0):
          kill move_thread_han_1745
          stopl(0.5)
          $ 1746 "Until (tool_contact_detection)"
          break
        end
        sleep(1.0E-10)
        if (move_thread_flag_1745 > 1):
          join move_thread_han_1745
          break
        end
        sync()
      end
      $ 1747 "Force"
      sleep(0.02)
      zero_ftsensor()
      force_mode(FRM_Reference, [1, 1, 1, 0, 0, 0], [0.0, 0.0, 0.0, 0.0, 0.0, 0.0], 2, [0.1, 0.1, 0.01, 0.3490658503988659, 0.3490658503988659, 0.3490658503988659])
      $ 1748 "PSE_T" "noBreak"
      movel(pose_trans(FRM_Reference, PSE_T), a=0.04, v=0.07)
      end_force_mode()
      stopl(5.0)
      $ 1749 "EXTT"
      $ 1750 "Switch JIG"
      switch_2 = JIG
      $ 1751 "Case 1"
      if (1 == switch_2):
        $ 1752 "3FG"
        $ 1753 "If OBJ_Picked"
        if (OBJ_Picked):
          $ 1754 "Set GRP_3F_Open=Off"
          set_standard_digital_out(5, False)
          $ 1755 "Wait: 0.2"
          sleep(0.2)
        end
      end
      $ 1756 "EOAT"
      $ 1757 "rq_move_and_wait_mm(GRP_Open_Pos)"
       rq_move_and_wait_mm (GRP_Open_Pos)
      $ 1758 "OBJ_Picked≔rq_is_object_detected()"
      global OBJ_Picked= rq_is_object_detected ()
      $ 1759 "If PSE_R_H≠PSE_Z"
      if (PSE_R_H != PSE_Z):
        $ 1760 "PSE_R" "breakAfter"
        movel(pose_trans(FRM_Reference, PSE_R), a=0.5, v=0.4, r=0.01)
        $ 1761 "PSE_R_H" "breakAfter"
        movel(pose_trans(FRM_Reference, PSE_R_H), a=0.5, v=0.4)
      else:
        $ 1762 "Else" "noBreak"
        $ 1763 "PSE_R" "breakAfter"
        movel(pose_trans(FRM_Reference, PSE_R), a=0.5, v=0.4)
      end
    elif (3 == switch_1):
      $ 1764 "Case 3"
      $ 1765 "Push"
      $ 1766 "Action_Info≔'push'"
      global Action_Info="push"
    elif (4 == switch_1):
      $ 1767 "Case 4"
      $ 1768 "Pull"
      $ 1769 "Action_Info≔'pull'"
      global Action_Info="pull"
    elif (6 == switch_1):
      $ 1772 "Case 6"
      $ 1773 "Drop the cap"
      $ 1774 "If JNT_A≠[0,0,0,0,0,0]"
      if (JNT_A != [0,0,0,0,0,0]):
        $ 1775 "MoveJ"
        $ 1776 "JNT_A" "breakAfter"
        movej(JNT_A, a=1.3962634015954636, v=1.7453292519943295, r=0.02)
      else:
        $ 1777 "Else" "noBreak"
        $ 1778 "MoveJ"
        $ 1779 "PSE_A" "breakAfter"
        movej(pose_trans(FRM_Reference, PSE_A), a=1.3962634015954636, v=1.7453292519943295, r=0.02)
      end
      $ 1780 "MoveL"
      $ 1781 "PSE_T" "breakAfter"
      movel(pose_trans(FRM_Reference, PSE_T), a=0.05, v=0.09)
      $ 1782 "'ADD OPEN GRIPPER'"
      # 'ADD OPEN GRIPPER'
      # begin: URCap Program Node
      #   Source: Robotiq_Grippers, 1.8.4.4844, Robotiq Inc.
      #   Type: Gripper
      $ 1783 "Gripper Move10mm (1)"
      if not(gripper_connected[0]):
        popup("Gripper 1 must be connected to run this program.", "No connection", False, True, True)
      end
      if not(rq_is_gripper_activated("1")):
        popup("Gripper 1 is not activated. Go to Installation tab > Gripper to activate it and run the program again.", "Not activated", False, True, True)
      end
      rq_set_pos_spd_for(201, 0, 28, "1")
      rq_wait_pos_spe_for_request(201, 0, 28, "1")
      rq_go_to("1")
      rq_wait("1")
      # end: URCap Program Node
      $ 1784 "PSE_T_H" "breakAfter"
      movel(pose_trans(FRM_Reference, PSE_T_H), a=0.05, v=0.09)
      # begin: URCap Program Node
      #   Source: Robotiq_Grippers, 1.8.4.4844, Robotiq Inc.
      #   Type: Gripper
      $ 1785 "Gripper Move40mm (1)"
      if not(gripper_connected[0]):
        popup("Gripper 1 must be connected to run this program.", "No connection", False, True, True)
      end
      if not(rq_is_gripper_activated("1")):
        popup("Gripper 1 is not activated. Go to Installation tab > Gripper to activate it and run the program again.", "Not activated", False, True, True)
      end
      rq_set_pos_spd_for(63, 0, 28, "1")
      rq_wait_pos_spe_for_request(63, 0, 28, "1")
      rq_go_to("1")
      rq_wait("1")
      # end: URCap Program Node
      $ 1786 "PSE_R" "breakAfter"
      movel(pose_trans(FRM_Reference, PSE_R), a=0.5, v=0.4)
    elif (7 == switch_1):
      $ 1787 "Case 7"
      $ 1788 "Load"
      $ 1789 "Action_Info≔'load object'"
      global Action_Info="load object"
      $ 1790 "do_transition(pose_trans(FRM_Reference, PSE_T), keep_rxry=OBJ_Picked)"
      do_transition( pose_trans (FRM_Reference, PSE_T), keep_rxry=OBJ_Picked)
      $ 1791 "If PSE_A_H≠PSE_Z"
      if (PSE_A_H != PSE_Z):
        $ 1792 "If JNT_Q≠JNT_Z"
        if (JNT_Q != JNT_Z):
          $ 1793 "movej(get_inverse_kin(pose_trans(FRM_Reference, PSE_A_H), qnear=JNT_Q), r=0.050)"
          movej(get_inverse_kin( pose_trans (FRM_Reference, PSE_A_H), qnear=JNT_Q), r=0.050)
        else:
          $ 1794 "Else" "noBreak"
          $ 1795 "movej(pose_trans(FRM_Reference, PSE_A_H), r=0.050)"
          movej( pose_trans (FRM_Reference, PSE_A_H), r=0.050)
        end
      end
      $ 1796 "If PSE_A≠PSE_Z"
      if (PSE_A != PSE_Z):
        $ 1797 "If JNT_Q≠JNT_Z"
        if (JNT_Q != JNT_Z):
          $ 1798 "movej(get_inverse_kin(pose_trans(FRM_Reference, PSE_A), qnear=JNT_Q), r=0.020)"
          movej(get_inverse_kin( pose_trans (FRM_Reference, PSE_A), qnear=JNT_Q), r=0.020)
        else:
          $ 1799 "Else" "noBreak"
          $ 1800 "movej(pose_trans(FRM_Reference, PSE_A), r=0.020)"
          movej( pose_trans (FRM_Reference, PSE_A), r=0.020)
        end
      end
      $ 1801 "MoveL"
      $ 1802 "If PSE_T_H≠PSE_Z"
      if (PSE_T_H != PSE_Z):
        $ 1803 "PSE_T_H" "breakAfter"
        movel(pose_trans(FRM_Reference, PSE_T_H), a=0.5, v=0.4, r=0.01)
      end
      $ 1804 "PSE_T" "breakAfter"
      global move_thread_flag_1804=0
      thread move_thread_1804():
        enter_critical
        move_thread_flag_1804 = 1
        movel(pose_trans(FRM_Reference, PSE_T), a=0.05, v=0.09)
        move_thread_flag_1804 = 2
        exit_critical
      end
      move_thread_flag_1804 = 0
      move_thread_han_1804 = run move_thread_1804()
      while (True):
        local targetTcpDirection=get_target_tcp_speed()
        local stepsToRetract=tool_contact(direction=targetTcpDirection)
        if (stepsToRetract > 0):
          kill move_thread_han_1804
          stopl(0.5)
          $ 1805 "Until (tool_contact_detection)"
          break
        end
        sleep(1.0E-10)
        if (move_thread_flag_1804 > 1):
          join move_thread_han_1804
          break
        end
        sync()
      end
      $ 1806 "Force"
      sleep(0.02)
      zero_ftsensor()
      force_mode(FRM_Reference, [0, 1, 1, 0, 0, 1], [0.0, 0.0, 0.0, 0.0, 0.0, 0.0], 2, [0.1, 0.05, 0.02, 0.3490658503988659, 0.3490658503988659, 3.141592653589793])
      $ 1807 "PSE_T" "noBreak"
      movel(pose_trans(FRM_Reference, PSE_T), a=0.04, v=0.07)
      end_force_mode()
      stopl(5.0)
      $ 1808 "EOAT"
      $ 1809 "rq_move_and_wait_mm(GRP_Open_Pos)"
       rq_move_and_wait_mm (GRP_Open_Pos)
      $ 1810 "OBJ_Picked≔rq_is_object_detected()"
      global OBJ_Picked= rq_is_object_detected ()
      $ 1811 "If PSE_R_H≠PSE_Z"
      if (PSE_R_H != PSE_Z):
        $ 1812 "PSE_R" "breakAfter"
        movel(pose_trans(FRM_Reference, PSE_R), a=0.5, v=0.4, r=0.01)
        $ 1813 "PSE_R_H" "breakAfter"
        movel(pose_trans(FRM_Reference, PSE_R_H), a=0.5, v=0.4)
      else:
        $ 1814 "Else" "noBreak"
        $ 1815 "PSE_R" "breakAfter"
        movel(pose_trans(FRM_Reference, PSE_R), a=0.5, v=0.4)
      end
    elif (8 == switch_1):
      $ 1816 "Case 8"
      $ 1817 "Unload"
      $ 1818 "Action_Info≔'pick object'"
      global Action_Info="pick object"
      $ 1819 "do_transition(pose_trans(FRM_Reference, PSE_T), keep_rxry=OBJ_Picked)"
      do_transition( pose_trans (FRM_Reference, PSE_T), keep_rxry=OBJ_Picked)
      $ 1820 "EOAT"
      $ 1821 "If  not OBJ_Picked"
      if (  not  OBJ_Picked):
        $ 1822 "rq_move_and_wait_mm(GRP_Open_Pos)"
         rq_move_and_wait_mm (GRP_Open_Pos)
      end
      $ 1823 "If PSE_A_H≠PSE_Z"
      if (PSE_A_H != PSE_Z):
        $ 1824 "If JNT_Q≠JNT_Z"
        if (JNT_Q != JNT_Z):
          $ 1825 "movej(get_inverse_kin(pose_trans(FRM_Reference, PSE_A_H), qnear=JNT_Q), r=0.050)"
          movej(get_inverse_kin( pose_trans (FRM_Reference, PSE_A_H), qnear=JNT_Q), r=0.050)
        else:
          $ 1826 "Else" "noBreak"
          $ 1827 "movej(pose_trans(FRM_Reference, PSE_A_H), r=0.050)"
          movej( pose_trans (FRM_Reference, PSE_A_H), r=0.050)
        end
      end
      $ 1828 "If PSE_A≠PSE_Z"
      if (PSE_A != PSE_Z):
        $ 1829 "If JNT_Q≠JNT_Z"
        if (JNT_Q != JNT_Z):
          $ 1830 "movej(get_inverse_kin(pose_trans(FRM_Reference, PSE_A), qnear=JNT_Q), r=0.020)"
          movej(get_inverse_kin( pose_trans (FRM_Reference, PSE_A), qnear=JNT_Q), r=0.020)
        else:
          $ 1831 "Else" "noBreak"
          $ 1832 "movej(pose_trans(FRM_Reference, PSE_A), r=0.020)"
          movej( pose_trans (FRM_Reference, PSE_A), r=0.020)
        end
      end
      $ 1833 "MoveL"
      $ 1834 "If PSE_T_H≠PSE_Z"
      if (PSE_T_H != PSE_Z):
        $ 1835 "PSE_T_H" "breakAfter"
        movel(pose_trans(FRM_Reference, PSE_T_H), a=0.5, v=0.4, r=0.01)
      end
      $ 1836 "PSE_T" "breakAfter"
      movel(pose_trans(FRM_Reference, PSE_T), a=0.08, v=0.12)
      $ 1837 "Force"
      sleep(0.02)
      zero_ftsensor()
      force_mode(FRM_Reference, [1, 1, 0, 0, 0, 0], [0.0, 0.0, 0.0, 0.0, 0.0, 0.0], 2, [0.05, 0.05, 0.1, 0.3490658503988659, 0.3490658503988659, 0.3490658503988659])
      $ 1838 "EOAT" "noBreak"
      $ 1839 "rq_set_force_norm(50)" "noBreak"
       rq_set_force_norm (50)
      $ 1840 "rq_close_and_wait()" "noBreak"
       rq_close_and_wait ()
      $ 1841 "OBJ_Picked≔rq_is_object_detected()" "noBreak"
      global OBJ_Picked= rq_is_object_detected ()
      $ 1842 "If  not OBJ_Picked" "noBreak"
      if (  not  OBJ_Picked):
        $ 1843 "set_error(ERROR_NO_OBJECT_TO_PICK)" "noBreak"
        set_error(ERROR_NO_OBJECT_TO_PICK)
      end
      $ 1844 "If PSE_R_H≠PSE_Z" "noBreak"
      if (PSE_R_H != PSE_Z):
        $ 1845 "PSE_R" "noBreak"
        movel(pose_trans(FRM_Reference, PSE_R), a=0.5, v=0.4, r=0.01)
        $ 1846 "PSE_R_H" "noBreak"
        movel(pose_trans(FRM_Reference, PSE_R_H), a=0.5, v=0.4)
      else:
        $ 1847 "Else" "noBreak"
        $ 1848 "PSE_R" "noBreak"
        movel(pose_trans(FRM_Reference, PSE_R), a=0.5, v=0.4)
      end
      end_force_mode()
      stopl(5.0)
    elif (11 == switch_1):
      $ 1849 "Case 11"
      $ 1850 "Place without opening gripper"
      $ 1851 "Action_Info≔'place object without gripper opening'"
      global Action_Info="place object without gripper opening"
      $ 1852 "do_transition(pose_trans(FRM_Reference, PSE_T), keep_rxry=OBJ_Picked)"
      do_transition( pose_trans (FRM_Reference, PSE_T), keep_rxry=OBJ_Picked)
      $ 1853 "EXTT"
      $ 1854 "Switch JIG"
      switch_2 = JIG
      $ 1855 "Case 1"
      if (1 == switch_2):
        $ 1856 "3FG"
        $ 1857 "If OBJ_Picked"
        if (OBJ_Picked):
          $ 1858 "Set GRP_3F_Open=On"
          set_standard_digital_out(5, True)
        end
      end
      $ 1859 "If PSE_A_H≠PSE_Z"
      if (PSE_A_H != PSE_Z):
        $ 1860 "If JNT_Q≠JNT_Z"
        if (JNT_Q != JNT_Z):
          $ 1861 "movej(get_inverse_kin(pose_trans(FRM_Reference, PSE_A_H), qnear=JNT_Q), r=0.050)"
          movej(get_inverse_kin( pose_trans (FRM_Reference, PSE_A_H), qnear=JNT_Q), r=0.050)
        else:
          $ 1862 "Else" "noBreak"
          $ 1863 "movej(pose_trans(FRM_Reference, PSE_A_H), r=0.050)"
          movej( pose_trans (FRM_Reference, PSE_A_H), r=0.050)
        end
      end
      $ 1864 "If PSE_A≠PSE_Z"
      if (PSE_A != PSE_Z):
        $ 1865 "If JNT_Q≠JNT_Z"
        if (JNT_Q != JNT_Z):
          $ 1866 "movej(get_inverse_kin(pose_trans(FRM_Reference, PSE_A), qnear=JNT_Q), r=0.020)"
          movej(get_inverse_kin( pose_trans (FRM_Reference, PSE_A), qnear=JNT_Q), r=0.020)
        else:
          $ 1867 "Else" "noBreak"
          $ 1868 "movej(pose_trans(FRM_Reference, PSE_A), r=0.020)"
          movej( pose_trans (FRM_Reference, PSE_A), r=0.020)
        end
      end
      $ 1869 "MoveL"
      $ 1870 "If PSE_T_H≠PSE_Z"
      if (PSE_T_H != PSE_Z):
        $ 1871 "PSE_T_H" "breakAfter"
        movel(pose_trans(FRM_Reference, PSE_T_H), a=0.5, v=0.4, r=0.01)
      end
      $ 1872 "PSE_T" "breakAfter"
      global move_thread_flag_1872=0
      thread move_thread_1872():
        enter_critical
        move_thread_flag_1872 = 1
        movel(pose_trans(FRM_Reference, PSE_T), a=0.05, v=0.09)
        move_thread_flag_1872 = 2
        exit_critical
      end
      move_thread_flag_1872 = 0
      move_thread_han_1872 = run move_thread_1872()
      while (True):
        local targetTcpDirection=get_target_tcp_speed()
        local stepsToRetract=tool_contact(direction=targetTcpDirection)
        if (stepsToRetract > 0):
          kill move_thread_han_1872
          stopl(0.5)
          $ 1873 "Until (tool_contact_detection)"
          break
        end
        sleep(1.0E-10)
        if (move_thread_flag_1872 > 1):
          join move_thread_han_1872
          break
        end
        sync()
      end
      $ 1874 "Force"
      sleep(0.02)
      zero_ftsensor()
      force_mode(FRM_Reference, [1, 1, 1, 0, 0, 0], [0.0, 0.0, 0.0, 0.0, 0.0, 0.0], 2, [0.1, 0.1, 0.01, 0.3490658503988659, 0.3490658503988659, 0.3490658503988659])
      $ 1875 "PSE_T" "noBreak"
      movel(pose_trans(FRM_Reference, PSE_T), a=0.04, v=0.07)
      end_force_mode()
      stopl(5.0)
      $ 1876 "EXTT"
      $ 1877 "Switch JIG"
      switch_2 = JIG
      $ 1878 "Case 1"
      if (1 == switch_2):
        $ 1879 "3FG"
        $ 1880 "If OBJ_Picked"
        if (OBJ_Picked):
          $ 1881 "Set GRP_3F_Open=Off"
          set_standard_digital_out(5, False)
          $ 1882 "Wait: 0.2"
          sleep(0.2)
        end
      end
      $ 1883 "EOAT"
      $ 1884 "Comment"
      # Comment
    elif (12 == switch_1):
      $ 1885 "Case 12"
      $ 1886 "Decap"
      $ 1887 "Action_Info≔'decapping'"
      global Action_Info="decapping"
      $ 1888 "Set GRP_3F_Enable=On"
      set_standard_digital_out(4, True)
      $ 1889 "Set GRP_3F_Decap=On"
      set_standard_digital_out(3, True)
      $ 1890 "Force"
      sleep(0.02)
      zero_ftsensor()
      force_mode(tool_pose(), [0, 0, 1, 0, 0, 0], [0.0, 0.0, 5.0, 0.0, 0.0, 0.0], 2, [0.1, 0.1, 0.15, 0.3490658503988659, 0.3490658503988659, 0.3490658503988659])
      $ 1891 "check_decapping(offset=0.015, timeout=5, abort=CMD_Hold)" "noBreak"
      check_decapping(offset=0.015, timeout=5, abort=CMD_Hold)
      end_force_mode()
      stopl(5.0)
      $ 1892 "Set GRP_3F_Decap=Off"
      set_standard_digital_out(3, False)
      $ 1893 "Set GRP_3F_Enable=Off"
      set_standard_digital_out(4, False)
      $ 1894 "MoveL"
      $ 1895 "PSE_R" "breakAfter"
      movel(pose_trans(FRM_Reference, PSE_R), a=0.8, v=0.15)
    elif (13 == switch_1):
      $ 1896 "Case 13"
      $ 1897 "TMR_Barcode: Reset"
      TMR_Barcode = 0
      $ 1898 "Read"
      $ 1899 "TMR_Barcode: Start"
      TMR_Barcode_is_counting = True
      $ 1900 "If TMR_Barcode<PRM_TO_Read_BC"
      global thread_flag_1900=0
      thread Thread_if_1900():
        $ 1901 "KeyenceTrigger"
        $ 1902 "Set OClearResult=HI:Pulse 0.2"
        thread SinglePulse88():
          write_output_boolean_register(2, True)
          sleep(0.2)
          write_output_boolean_register(2, False)
        end
        singlePulse88 = run SinglePulse88()
        $ 1903 "Wait: 0.5"
        sleep(0.5)
        $ 1904 "Set OTriggerBarcode=Off"
        write_output_boolean_register(1, False)
        $ 1905 "Wait: 0.5"
        sleep(0.5)
        $ 1906 "Set OTriggerBarcode=On"
        write_output_boolean_register(1, True)
        $ 1907 "Wait: 0.5"
        sleep(0.5)
        $ 1908 "Preorient"
        $ 1909 "TMR_Barcode: Reset"
        TMR_Barcode = 0
        $ 1910 "If ICmdExctd"
        if (read_input_boolean_register(12)):
          $ 1911 "Set GRP_3F_Decap=On"
          set_standard_digital_out(3, True)
          $ 1912 "Set GRP_3F_Enable=On"
          set_standard_digital_out(4, True)
          $ 1913 "Loop ICmdExctd"
          while (read_input_boolean_register(12)):
            $ 1914 "KeyenceTrigger"
            $ 1915 "Set OClearResult=HI:Pulse 0.1"
            thread SinglePulse89():
              write_output_boolean_register(2, True)
              sleep(0.1)
              write_output_boolean_register(2, False)
            end
            singlePulse89 = run SinglePulse89()
            $ 1916 "Wait: 0.3"
            sleep(0.3)
            $ 1917 "Set OTriggerBarcode=Off"
            write_output_boolean_register(1, False)
            $ 1918 "Wait: 0.3"
            sleep(0.3)
            $ 1919 "Set OTriggerBarcode=On"
            write_output_boolean_register(1, True)
            $ 1920 "Wait: 0.1"
            sleep(0.1)
          end
        end
        $ 1921 "If  not ICmdExctd"
        if (  not  read_input_boolean_register(12)):
          $ 1922 "Set GRP_3F_Decap=On"
          set_standard_digital_out(3, True)
          $ 1923 "Set GRP_3F_Enable=On"
          set_standard_digital_out(4, True)
          $ 1924 "Wait ICmdExctd=HI"
          while (read_input_boolean_register(12) == False):
            sync()
          end
        end
        $ 1925 "Set GRP_3F_Decap=Off"
        set_standard_digital_out(3, False)
        $ 1926 "Set GRP_3F_Enable=Off"
        set_standard_digital_out(4, False)
        $ 1927 "OBJ_Brc_OK≔ True "
        global OBJ_Brc_OK=  True
        thread_flag_1900 = 1
      end
      if (TMR_Barcode<PRM_TO_Read_BC):
        global thread_handler_1900=run Thread_if_1900()
        while (thread_flag_1900 == 0):
          if not(TMR_Barcode<PRM_TO_Read_BC):
            kill thread_handler_1900
            thread_flag_1900 = 2
          else:
            sync()
          end
        end
      else:
        thread_flag_1900 = 2
      end
      if (thread_flag_1900 == 2):
        $ 1928 "Else" "noBreak"
        $ 1929 "exeption"
        $ 1930 "error"
        $ 1932 "OBJ_Brc_OK≔ False "
        global OBJ_Brc_OK=  False
      end
      $ 1933 "Set GRP_3F_Decap=Off"
      set_standard_digital_out(3, False)
      $ 1934 "Set GRP_3F_Enable=Off"
      set_standard_digital_out(4, False)
      $ 1935 "Set OTriggerBarcode=Off"
      write_output_boolean_register(1, False)
    elif (15 == switch_1):
      $ 1936 "Case 15"
      $ 1937 "Detect"
      $ 1938 "Action_Info≔'detect'"
      global Action_Info="detect"
    elif (30 == switch_1):
      $ 1939 "Case 30"
      $ 1940 "Shake"
      $ 1941 "Action_Info≔'shake'"
      global Action_Info="shake"
      $ 1942 "do_transition(pose_trans(FRM_Reference, PSE_T), keep_rxry=OBJ_Picked)"
      do_transition( pose_trans (FRM_Reference, PSE_T), keep_rxry=OBJ_Picked)
      $ 1943 "If PSE_A_H≠PSE_Z"
      if (PSE_A_H != PSE_Z):
        $ 1944 "If JNT_Q≠JNT_Z"
        if (JNT_Q != JNT_Z):
          $ 1945 "movej(get_inverse_kin(pose_trans(FRM_Reference, PSE_A_H), qnear=JNT_Q), r=0.050)"
          movej(get_inverse_kin( pose_trans (FRM_Reference, PSE_A_H), qnear=JNT_Q), r=0.050)
        else:
          $ 1946 "Else" "noBreak"
          $ 1947 "movej(pose_trans(FRM_Reference, PSE_A_H), r=0.050)"
          movej( pose_trans (FRM_Reference, PSE_A_H), r=0.050)
        end
      end
      $ 1948 "If PSE_A≠PSE_Z"
      if (PSE_A != PSE_Z):
        $ 1949 "If JNT_Q≠JNT_Z"
        if (JNT_Q != JNT_Z):
          $ 1950 "movej(get_inverse_kin(pose_trans(FRM_Reference, PSE_A), qnear=JNT_Q), r=0.020)"
          movej(get_inverse_kin( pose_trans (FRM_Reference, PSE_A), qnear=JNT_Q), r=0.020)
        else:
          $ 1951 "Else" "noBreak"
          $ 1952 "movej(pose_trans(FRM_Reference, PSE_A), r=0.020)"
          movej( pose_trans (FRM_Reference, PSE_A), r=0.020)
        end
      end
      $ 1953 "MoveL"
      $ 1954 "If PSE_T_H≠PSE_Z"
      if (PSE_T_H != PSE_Z):
        $ 1955 "PSE_T_H" "breakAfter"
        movel(pose_trans(FRM_Reference, PSE_T_H), a=0.5, v=0.4, r=0.01)
      end
      $ 1956 "PSE_T" "breakAfter"
      movel(pose_trans(FRM_Reference, PSE_T), a=0.08, v=0.12)
      $ 1957 "EXTT"
      $ 1958 "Comment"
      # Comment
      $ 1959 "MoveJ"
      $ 1960 "Waypoint_6" "breakAfter"
      movej(get_inverse_kin(Waypoint_6_p, qnear=Waypoint_6_q), a=1.3962634015954636, v=1.0471975511965976)
      $ 1961 "MoveJ"
      $ 1962 "Waypoint_18" "breakAfter"
      movej(get_inverse_kin(Waypoint_18_p, qnear=Waypoint_18_q), a=1.3962634015954636, v=1.0471975511965976)
      $ 1963 "MoveJ"
      $ 1964 "Waypoint_12" "breakAfter"
      movej(get_inverse_kin(Waypoint_12_p, qnear=Waypoint_12_q), a=1.3962634015954636, v=1.0471975511965976)
      $ 1965 "MoveJ"
      $ 1966 "Waypoint_19" "breakAfter"
      movej(get_inverse_kin(Waypoint_19_p, qnear=Waypoint_19_q), a=1.3962634015954636, v=1.0471975511965976)
      $ 1967 "If PSE_R_H≠PSE_Z"
      if (PSE_R_H != PSE_Z):
        $ 1968 "PSE_R" "breakAfter"
        movel(pose_trans(FRM_Reference, PSE_R), a=0.5, v=0.4, r=0.01)
        $ 1969 "PSE_R_H" "breakAfter"
        movel(pose_trans(FRM_Reference, PSE_R_H), a=0.5, v=0.4)
      else:
        $ 1970 "Else" "noBreak"
        $ 1971 "PSE_R" "breakAfter"
        movel(pose_trans(FRM_Reference, PSE_R), a=0.5, v=0.4)
      end
    elif (31 == switch_1):
      $ 1972 "Case 31"
      $ 1973 "Action_Info≔'Pick_Vial'"
      global Action_Info="Pick_Vial"
      $ 1974 "Pick_Vial"
      # begin: URCap Program Node
      #   Source: Robotiq_Grippers, 1.8.4.4844, Robotiq Inc.
      #   Type: Gripper
      $ 1975 "Gripper Open (1)"
      if not(gripper_connected[0]):
        popup("Gripper 1 must be connected to run this program.", "No connection", False, True, True)
      end
      if not(rq_is_gripper_activated("1")):
        popup("Gripper 1 is not activated. Go to Installation tab > Gripper to activate it and run the program again.", "Not activated", False, True, True)
      end
      rq_set_pos_spd_for(0, 82, 71, "1")
      rq_wait_pos_spe_for_request(0, 82, 71, "1")
      rq_go_to("1")
      rq_wait("1")
      # end: URCap Program Node
      $ 1976 "MoveJ"
      $ 1977 "Vial_above" "breakAfter"
      movej(get_inverse_kin(Vial_above_p, qnear=Vial_above_q), a=0.5235987755982988, v=0.4363323129985824, r=0.05)
      $ 1978 "MoveL"
      $ 1979 "Vial_pick_point" "breakAfter"
      movel(Vial_pick_point_p, a=0.5, v=0.1)
      # begin: URCap Program Node
      #   Source: Robotiq_Grippers, 1.8.4.4844, Robotiq Inc.
      #   Type: Gripper
      $ 1980 "Gripper Close (1)"
      if not(gripper_connected[0]):
        popup("Gripper 1 must be connected to run this program.", "No connection", False, True, True)
      end
      if not(rq_is_gripper_activated("1")):
        popup("Gripper 1 is not activated. Go to Installation tab > Gripper to activate it and run the program again.", "Not activated", False, True, True)
      end
      rq_set_pos_spd_for(255, 71, 84, "1")
      rq_wait_pos_spe_for_request(255, 71, 84, "1")
      rq_go_to("1")
      rq_wait("1")
      # end: URCap Program Node
      $ 1981 "MoveL"
      $ 1982 "Waypoint_20" "breakAfter"
      movel(Waypoint_20_p, a=0.5, v=0.1, r=0.05)
      $ 1983 "Home (Safe)"
      movej([-1.2302089344500047, -1.2969853503591224, -1.875639182904262, -1.539621866126728, 1.5731943360401213, -2.80099559440227], a=1.3962634015954636, v=1.0471975511965976)
    elif (32 == switch_1):
      $ 1984 "Case 32"
      $ 1985 "decap≔ False "
      global decap=  False
      $ 1986 "decap_Vial"
      $ 1987 "Set GRP_3F_Open=On"
      set_standard_digital_out(5, True)
      $ 1988 "MoveJ"
      $ 1989 "Waypoint_33" "breakAfter"
      movej(get_inverse_kin(Waypoint_33_p, qnear=Waypoint_33_q), a=0.5235987755982988, v=0.4363323129985824)
      $ 1990 "MoveL"
      $ 1991 "Vial_3FG_place" "breakAfter"
      movel(Vial_3FG_place_p, a=0.5, v=0.1)
      $ 1992 "Set GRP_3F_Open=Off"
      set_standard_digital_out(5, False)
      $ 1993 "Wait: 0.5"
      sleep(0.5)
      $ 1994 "MoveL"
      $ 1995 "Waypoint_34" "breakAfter"
      movel(Waypoint_34_p, a=0.5, v=0.1, r=0.05)
      $ 1996 "MoveJ"
      $ 1997 "cap_dump" "breakAfter"
      movej(get_inverse_kin(cap_dump_p, qnear=cap_dump_q), a=0.5235987755982988, v=0.4363323129985824)
      # begin: URCap Program Node
      #   Source: Robotiq_Grippers, 1.8.4.4844, Robotiq Inc.
      #   Type: Gripper
      $ 1998 "Gripper Open (1)"
      if not(gripper_connected[0]):
        popup("Gripper 1 must be connected to run this program.", "No connection", False, True, True)
      end
      if not(rq_is_gripper_activated("1")):
        popup("Gripper 1 is not activated. Go to Installation tab > Gripper to activate it and run the program again.", "Not activated", False, True, True)
      end
      rq_set_pos_spd_for(0, 255, 255, "1")
      rq_wait_pos_spe_for_request(0, 255, 255, "1")
      rq_go_to("1")
      rq_wait("1")
      # end: URCap Program Node
      $ 1999 "MoveJ"
      $ 2000 "Waypoint_35" "breakAfter"
      movej(get_inverse_kin(Waypoint_35_p, qnear=Waypoint_35_q), a=0.5235987755982988, v=0.4363323129985824, r=0.05)
      $ 2001 "MoveL"
      $ 2002 "Vial_3FG_place" "breakAfter"
      movel(Vial_3FG_place_p, a=0.5, v=0.1)
      # begin: URCap Program Node
